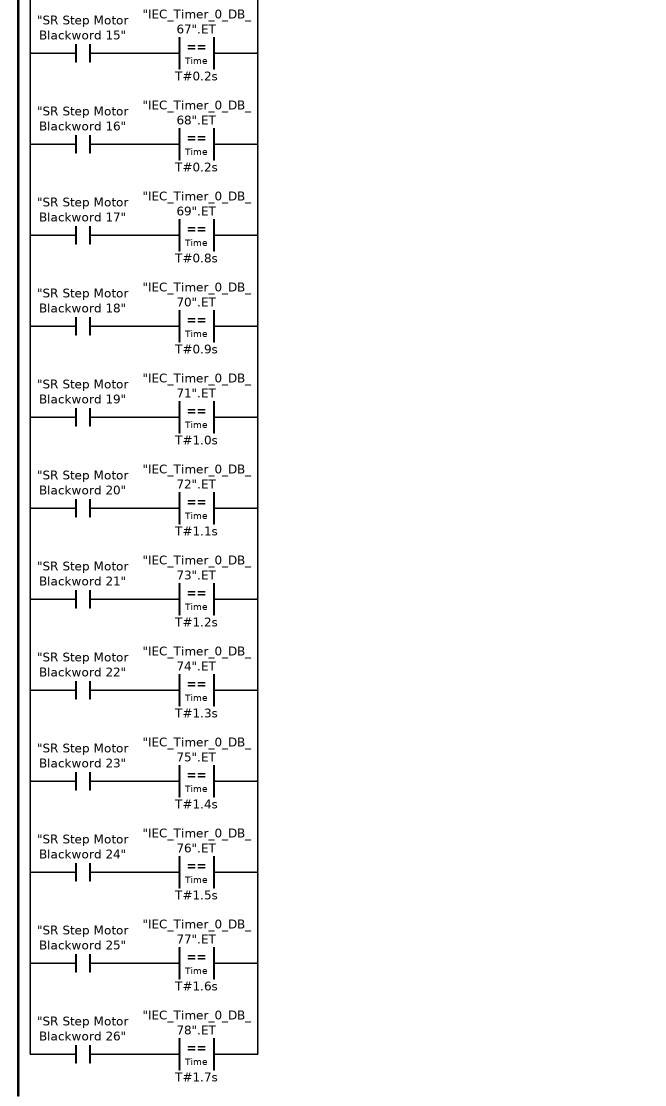
   "IEC_Counter_0_DB_1072".CTU(CU := ("SR Step Motor Blackword 1" AND ("IEC_Timer_0_DB_36".ET = T#2.0s)) OR ("SR Step Motor Blackword 2" AND ("IEC_Timer_0_DB_54".ET = T#1.9s)) OR ("SR Step Motor Blackword 3" AND ("IEC_Timer_0_DB_55".ET = T#1.8s)) OR ("SR Step Motor Blackword 4" AND ("IEC_Timer_0_DB_56".ET = T#1.7s)) OR ("SR Step Motor Blackword 5" AND ("IEC_Timer_0_DB_57".ET = T#1.6s)) OR ("SR Step Motor Blackword 6" AND ("IEC_Timer_0_DB_58".ET = T#1.5s)) OR ("SR Step Motor Blackword 7" AND ("IEC_Timer_0_DB_59".ET = T#1.4s)) OR ("SR Step Motor Blackword 8" AND ("IEC_Timer_0_DB_60".ET = T#1.3s)) OR ("SR Step Motor Blackword 9" AND ("IEC_Timer_0_DB_61".ET = T#1.2s)) OR ("SR Step Motor Blackword 10" AND ("IEC_Timer_0_DB_62".ET = T#1.1s)) OR ("SR Step Motor Blackword 11" AND ("IEC_Timer_0_DB_63".ET = T#1.0s)) OR ("SR Step Motor Blackword 12" AND ("IEC_Timer_0_DB_64".ET = T#0.9s)) OR ("SR Step Motor Blackword 13" AND ("IEC_Timer_0_DB_65".ET = T#0.8s)) OR ("SR Step Motor Blackword 14" AND ("IEC_Timer_0_DB_66".ET = T#0.2s)) OR ("SR Step Motor Blackword 15" AND ("IEC_Timer_0_DB_67".ET = T#0.2s)) OR ("SR Step Motor Blackword 16" AND ("IEC_Timer_0_DB_68".ET = T#0.2s)) OR ("SR Step Motor Blackword 17" AND ("IEC_Timer_0_DB_69".ET = T#0.8s)) OR ("SR Step Motor Blackword 18" AND ("IEC_Timer_0_DB_70".ET = T#0.9s)) OR ("SR Step Motor Blackword 19" AND ("IEC_Timer_0_DB_71".ET = T#1.0s)) OR ("SR Step Motor Blackword 20" AND ("IEC_Timer_0_DB_72".ET = T#1.1s)) OR ("SR Step Motor Blackword 21" AND ("IEC_Timer_0_DB_73".ET = T#1.2s)) OR ("SR Step Motor Blackword 22" AND ("IEC_Timer_0_DB_74".ET = T#1.3s)) OR ("SR Step Motor Blackword 23" AND ("IEC_Timer_0_DB_75".ET = T#1.4s)) OR ("SR Step Motor Blackword 24" AND ("IEC_Timer_0_DB_76".ET = T#1.5s)) OR ("SR Step Motor Blackword 25" AND ("IEC_Timer_0_DB_77".ET = T#1.6s)) OR ("SR Step Motor Blackword 26" AND ("IEC_Timer_0_DB_78".ET = T#1.7s)),
                           R := "Brushless Motor Conveyor ทำงาน",
                           PV := 1);
   "Output Reset พิเศษ จัดเก็บบ" := "IEC_Counter_0_DB_1072".Q;
END_REGION
END_FUNCTION_BLOCK

FUNCTION "Test" : Void   // FC5, LAD
{ S7_Optimized_Access := 'TRUE' }
VERSION : 0.1
BEGIN

REGION Network 1
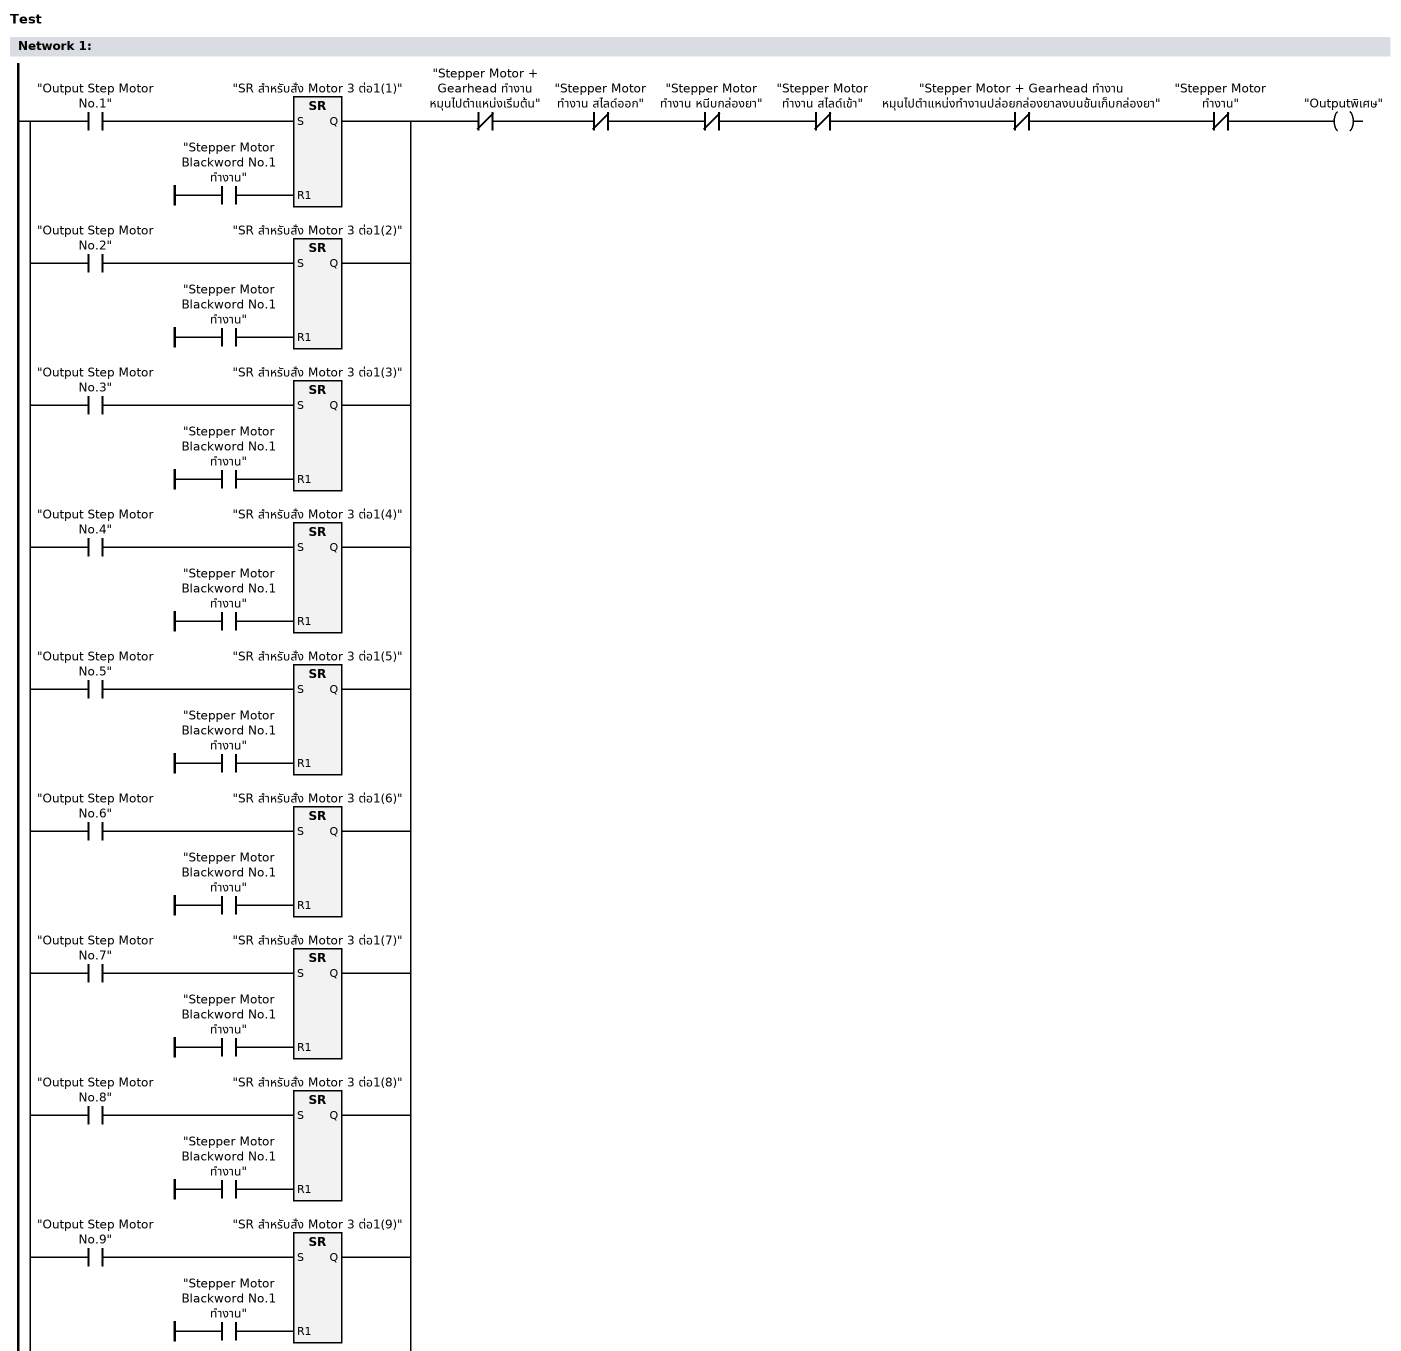
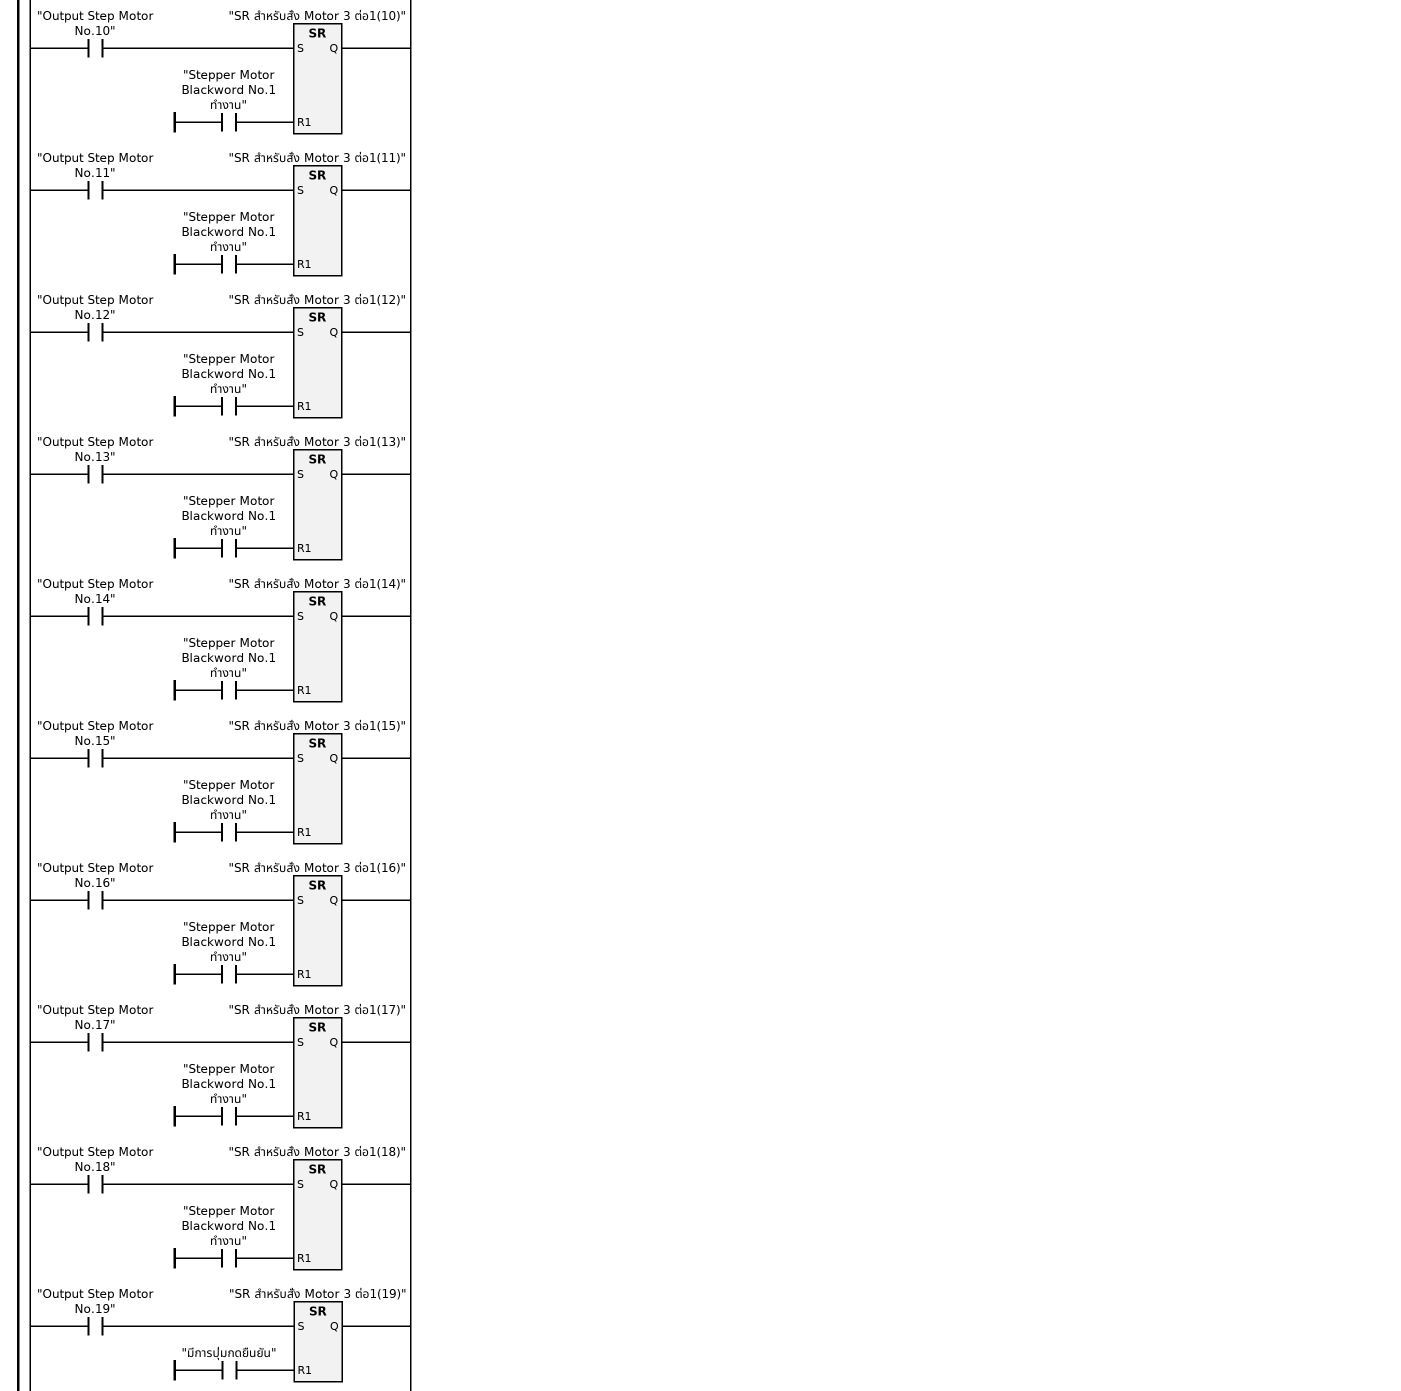
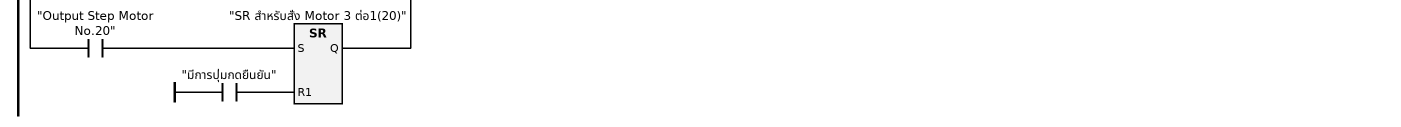
   RUNG wire#powerrail
      Contact( "Output Step Motor No.1" )
      S_SR(operand := "SR สำหรับสั่ง Motor 3 ต่อ1(1)", r1 := wire#w1)
      wire#w2
      I_Contact( "Stepper Motor + Gearhead ทำงาน หมุนไปตำแหน่งเริ่มต้น" )
      I_Contact( "Stepper Motor ทำงาน สไลด์ออก" )
      I_Contact( "Stepper Motor ทำงาน หนีบกล่องยา" )
      I_Contact( "Stepper Motor ทำงาน สไลด์เข้า" )
      I_Contact( "Stepper Motor + Gearhead ทำงาน หมุนไปตำแหน่งทำงานปล่อยกล่องยาลงบนชั้นเก็บกล่องยา" )
      I_Contact( "Stepper Motor  ทำงาน" )
      Coil( "Outputพิเศษ" )
   END_RUNG
   RUNG wire#powerrail
      Contact( "Stepper Motor Blackword No.1 ทำงาน" )
   END_RUNG wire#w1
   RUNG wire#powerrail
      Contact( "Output Step Motor No.2" )
      S_SR(operand := "SR สำหรับสั่ง Motor 3 ต่อ1(2)", r1 := wire#w3)
   END_RUNG wire#w2
   RUNG wire#powerrail
      Contact( "Stepper Motor Blackword No.1 ทำงาน" )
   END_RUNG wire#w3
   RUNG wire#powerrail
      Contact( "Output Step Motor No.3" )
      S_SR(operand := "SR สำหรับสั่ง Motor 3 ต่อ1(3)", r1 := wire#w4)
   END_RUNG wire#w2
   RUNG wire#powerrail
      Contact( "Stepper Motor Blackword No.1 ทำงาน" )
   END_RUNG wire#w4
   RUNG wire#powerrail
      Contact( "Output Step Motor No.4" )
      S_SR(operand := "SR สำหรับสั่ง Motor 3 ต่อ1(4)", r1 := wire#w5)
   END_RUNG wire#w2
   RUNG wire#powerrail
      Contact( "Stepper Motor Blackword No.1 ทำงาน" )
   END_RUNG wire#w5
   RUNG wire#powerrail
      Contact( "Output Step Motor No.5" )
      S_SR(operand := "SR สำหรับสั่ง Motor 3 ต่อ1(5)", r1 := wire#w6)
   END_RUNG wire#w2
   RUNG wire#powerrail
      Contact( "Stepper Motor Blackword No.1 ทำงาน" )
   END_RUNG wire#w6
   RUNG wire#powerrail
      Contact( "Output Step Motor No.6" )
      S_SR(operand := "SR สำหรับสั่ง Motor 3 ต่อ1(6)", r1 := wire#w7)
   END_RUNG wire#w2
   RUNG wire#powerrail
      Contact( "Stepper Motor Blackword No.1 ทำงาน" )
   END_RUNG wire#w7
   RUNG wire#powerrail
      Contact( "Output Step Motor No.7" )
      S_SR(operand := "SR สำหรับสั่ง Motor 3 ต่อ1(7)", r1 := wire#w8)
   END_RUNG wire#w2
   RUNG wire#powerrail
      Contact( "Stepper Motor Blackword No.1 ทำงาน" )
   END_RUNG wire#w8
   RUNG wire#powerrail
      Contact( "Output Step Motor No.8" )
      S_SR(operand := "SR สำหรับสั่ง Motor 3 ต่อ1(8)", r1 := wire#w9)
   END_RUNG wire#w2
   RUNG wire#powerrail
      Contact( "Stepper Motor Blackword No.1 ทำงาน" )
   END_RUNG wire#w9
   RUNG wire#powerrail
      Contact( "Output Step Motor No.9" )
      S_SR(operand := "SR สำหรับสั่ง Motor 3 ต่อ1(9)", r1 := wire#w10)
   END_RUNG wire#w2
   RUNG wire#powerrail
      Contact( "Stepper Motor Blackword No.1 ทำงาน" )
   END_RUNG wire#w10
   RUNG wire#powerrail
      Contact( "Output Step Motor No.10" )
      S_SR(operand := "SR สำหรับสั่ง Motor 3 ต่อ1(10)", r1 := wire#w11)
   END_RUNG wire#w2
   RUNG wire#powerrail
      Contact( "Stepper Motor Blackword No.1 ทำงาน" )
   END_RUNG wire#w11
   RUNG wire#powerrail
      Contact( "Output Step Motor No.11" )
      S_SR(operand := "SR สำหรับสั่ง Motor 3 ต่อ1(11)", r1 := wire#w12)
   END_RUNG wire#w2
   RUNG wire#powerrail
      Contact( "Stepper Motor Blackword No.1 ทำงาน" )
   END_RUNG wire#w12
   RUNG wire#powerrail
      Contact( "Output Step Motor No.12" )
      S_SR(operand := "SR สำหรับสั่ง Motor 3 ต่อ1(12)", r1 := wire#w13)
   END_RUNG wire#w2
   RUNG wire#powerrail
      Contact( "Stepper Motor Blackword No.1 ทำงาน" )
   END_RUNG wire#w13
   RUNG wire#powerrail
      Contact( "Output Step Motor No.13" )
      S_SR(operand := "SR สำหรับสั่ง Motor 3 ต่อ1(13)", r1 := wire#w14)
   END_RUNG wire#w2
   RUNG wire#powerrail
      Contact( "Stepper Motor Blackword No.1 ทำงาน" )
   END_RUNG wire#w14
   RUNG wire#powerrail
      Contact( "Output Step Motor No.14" )
      S_SR(operand := "SR สำหรับสั่ง Motor 3 ต่อ1(14)", r1 := wire#w15)
   END_RUNG wire#w2
   RUNG wire#powerrail
      Contact( "Stepper Motor Blackword No.1 ทำงาน" )
   END_RUNG wire#w15
   RUNG wire#powerrail
      Contact( "Output Step Motor No.15" )
      S_SR(operand := "SR สำหรับสั่ง Motor 3 ต่อ1(15)", r1 := wire#w16)
   END_RUNG wire#w2
   RUNG wire#powerrail
      Contact( "Stepper Motor Blackword No.1 ทำงาน" )
   END_RUNG wire#w16
   RUNG wire#powerrail
      Contact( "Output Step Motor No.16" )
      S_SR(operand := "SR สำหรับสั่ง Motor 3 ต่อ1(16)", r1 := wire#w17)
   END_RUNG wire#w2
   RUNG wire#powerrail
      Contact( "Stepper Motor Blackword No.1 ทำงาน" )
   END_RUNG wire#w17
   RUNG wire#powerrail
      Contact( "Output Step Motor No.17" )
      S_SR(operand := "SR สำหรับสั่ง Motor 3 ต่อ1(17)", r1 := wire#w18)
   END_RUNG wire#w2
   RUNG wire#powerrail
      Contact( "Stepper Motor Blackword No.1 ทำงาน" )
   END_RUNG wire#w18
   RUNG wire#powerrail
      Contact( "Output Step Motor No.18" )
      S_SR(operand := "SR สำหรับสั่ง Motor 3 ต่อ1(18)", r1 := wire#w19)
   END_RUNG wire#w2
   RUNG wire#powerrail
      Contact( "Stepper Motor Blackword No.1 ทำงาน" )
   END_RUNG wire#w19
   RUNG wire#powerrail
      Contact( "Output Step Motor No.19" )
      S_SR(operand := "SR สำหรับสั่ง Motor 3 ต่อ1(19)", r1 := wire#w20)
   END_RUNG wire#w2
   RUNG wire#powerrail
      Contact( "มีการปุ่มกดยืนยัน" )
   END_RUNG wire#w20
   RUNG wire#powerrail
      Contact( "Output Step Motor No.20" )
      S_SR(operand := "SR สำหรับสั่ง Motor 3 ต่อ1(20)", r1 := wire#w21)
   END_RUNG wire#w2
   RUNG wire#powerrail
      Contact( "มีการปุ่มกดยืนยัน" )
   END_RUNG wire#w21
   // the same network as SCL:
   IF "Output Step Motor No.1" THEN
       "SR สำหรับสั่ง Motor 3 ต่อ1(1)" := TRUE;   // SR flip-flop
   END_IF;
   IF "Stepper Motor Blackword No.1 ทำงาน" THEN "SR สำหรับสั่ง Motor 3 ต่อ1(1)" := FALSE; END_IF;
   IF "Output Step Motor No.2" THEN
       "SR สำหรับสั่ง Motor 3 ต่อ1(2)" := TRUE;   // SR flip-flop
   END_IF;
   IF "Stepper Motor Blackword No.1 ทำงาน" THEN "SR สำหรับสั่ง Motor 3 ต่อ1(2)" := FALSE; END_IF;
   IF "Output Step Motor No.3" THEN
       "SR สำหรับสั่ง Motor 3 ต่อ1(3)" := TRUE;   // SR flip-flop
   END_IF;
   IF "Stepper Motor Blackword No.1 ทำงาน" THEN "SR สำหรับสั่ง Motor 3 ต่อ1(3)" := FALSE; END_IF;
   IF "Output Step Motor No.4" THEN
       "SR สำหรับสั่ง Motor 3 ต่อ1(4)" := TRUE;   // SR flip-flop
   END_IF;
   IF "Stepper Motor Blackword No.1 ทำงาน" THEN "SR สำหรับสั่ง Motor 3 ต่อ1(4)" := FALSE; END_IF;
   IF "Output Step Motor No.5" THEN
       "SR สำหรับสั่ง Motor 3 ต่อ1(5)" := TRUE;   // SR flip-flop
   END_IF;
   IF "Stepper Motor Blackword No.1 ทำงาน" THEN "SR สำหรับสั่ง Motor 3 ต่อ1(5)" := FALSE; END_IF;
   IF "Output Step Motor No.6" THEN
       "SR สำหรับสั่ง Motor 3 ต่อ1(6)" := TRUE;   // SR flip-flop
   END_IF;
   IF "Stepper Motor Blackword No.1 ทำงาน" THEN "SR สำหรับสั่ง Motor 3 ต่อ1(6)" := FALSE; END_IF;
   IF "Output Step Motor No.7" THEN
       "SR สำหรับสั่ง Motor 3 ต่อ1(7)" := TRUE;   // SR flip-flop
   END_IF;
   IF "Stepper Motor Blackword No.1 ทำงาน" THEN "SR สำหรับสั่ง Motor 3 ต่อ1(7)" := FALSE; END_IF;
   IF "Output Step Motor No.8" THEN
       "SR สำหรับสั่ง Motor 3 ต่อ1(8)" := TRUE;   // SR flip-flop
   END_IF;
   IF "Stepper Motor Blackword No.1 ทำงาน" THEN "SR สำหรับสั่ง Motor 3 ต่อ1(8)" := FALSE; END_IF;
   IF "Output Step Motor No.9" THEN
       "SR สำหรับสั่ง Motor 3 ต่อ1(9)" := TRUE;   // SR flip-flop
   END_IF;
   IF "Stepper Motor Blackword No.1 ทำงาน" THEN "SR สำหรับสั่ง Motor 3 ต่อ1(9)" := FALSE; END_IF;
   IF "Output Step Motor No.10" THEN
       "SR สำหรับสั่ง Motor 3 ต่อ1(10)" := TRUE;   // SR flip-flop
   END_IF;
   IF "Stepper Motor Blackword No.1 ทำงาน" THEN "SR สำหรับสั่ง Motor 3 ต่อ1(10)" := FALSE; END_IF;
   IF "Output Step Motor No.11" THEN
       "SR สำหรับสั่ง Motor 3 ต่อ1(11)" := TRUE;   // SR flip-flop
   END_IF;
   IF "Stepper Motor Blackword No.1 ทำงาน" THEN "SR สำหรับสั่ง Motor 3 ต่อ1(11)" := FALSE; END_IF;
   IF "Output Step Motor No.12" THEN
       "SR สำหรับสั่ง Motor 3 ต่อ1(12)" := TRUE;   // SR flip-flop
   END_IF;
   IF "Stepper Motor Blackword No.1 ทำงาน" THEN "SR สำหรับสั่ง Motor 3 ต่อ1(12)" := FALSE; END_IF;
   IF "Output Step Motor No.13" THEN
       "SR สำหรับสั่ง Motor 3 ต่อ1(13)" := TRUE;   // SR flip-flop
   END_IF;
   IF "Stepper Motor Blackword No.1 ทำงาน" THEN "SR สำหรับสั่ง Motor 3 ต่อ1(13)" := FALSE; END_IF;
   IF "Output Step Motor No.14" THEN
       "SR สำหรับสั่ง Motor 3 ต่อ1(14)" := TRUE;   // SR flip-flop
   END_IF;
   IF "Stepper Motor Blackword No.1 ทำงาน" THEN "SR สำหรับสั่ง Motor 3 ต่อ1(14)" := FALSE; END_IF;
   IF "Output Step Motor No.15" THEN
       "SR สำหรับสั่ง Motor 3 ต่อ1(15)" := TRUE;   // SR flip-flop
   END_IF;
   IF "Stepper Motor Blackword No.1 ทำงาน" THEN "SR สำหรับสั่ง Motor 3 ต่อ1(15)" := FALSE; END_IF;
   IF "Output Step Motor No.16" THEN
       "SR สำหรับสั่ง Motor 3 ต่อ1(16)" := TRUE;   // SR flip-flop
   END_IF;
   IF "Stepper Motor Blackword No.1 ทำงาน" THEN "SR สำหรับสั่ง Motor 3 ต่อ1(16)" := FALSE; END_IF;
   IF "Output Step Motor No.17" THEN
       "SR สำหรับสั่ง Motor 3 ต่อ1(17)" := TRUE;   // SR flip-flop
   END_IF;
   IF "Stepper Motor Blackword No.1 ทำงาน" THEN "SR สำหรับสั่ง Motor 3 ต่อ1(17)" := FALSE; END_IF;
   IF "Output Step Motor No.18" THEN
       "SR สำหรับสั่ง Motor 3 ต่อ1(18)" := TRUE;   // SR flip-flop
   END_IF;
   IF "Stepper Motor Blackword No.1 ทำงาน" THEN "SR สำหรับสั่ง Motor 3 ต่อ1(18)" := FALSE; END_IF;
   IF "Output Step Motor No.19" THEN
       "SR สำหรับสั่ง Motor 3 ต่อ1(19)" := TRUE;   // SR flip-flop
   END_IF;
   IF "มีการปุ่มกดยืนยัน" THEN "SR สำหรับสั่ง Motor 3 ต่อ1(19)" := FALSE; END_IF;
   IF "Output Step Motor No.20" THEN
       "SR สำหรับสั่ง Motor 3 ต่อ1(20)" := TRUE;   // SR flip-flop
   END_IF;
   IF "มีการปุ่มกดยืนยัน" THEN "SR สำหรับสั่ง Motor 3 ต่อ1(20)" := FALSE; END_IF;
   "Outputพิเศษ" := ("SR สำหรับสั่ง Motor 3 ต่อ1(1)" OR "SR สำหรับสั่ง Motor 3 ต่อ1(2)" OR "SR สำหรับสั่ง Motor 3 ต่อ1(3)" OR "SR สำหรับสั่ง Motor 3 ต่อ1(4)" OR "SR สำหรับสั่ง Motor 3 ต่อ1(5)" OR "SR สำหรับสั่ง Motor 3 ต่อ1(6)" OR "SR สำหรับสั่ง Motor 3 ต่อ1(7)" OR "SR สำหรับสั่ง Motor 3 ต่อ1(8)" OR "SR สำหรับสั่ง Motor 3 ต่อ1(9)" OR "SR สำหรับสั่ง Motor 3 ต่อ1(10)" OR "SR สำหรับสั่ง Motor 3 ต่อ1(11)" OR "SR สำหรับสั่ง Motor 3 ต่อ1(12)" OR "SR สำหรับสั่ง Motor 3 ต่อ1(13)" OR "SR สำหรับสั่ง Motor 3 ต่อ1(14)" OR "SR สำหรับสั่ง Motor 3 ต่อ1(15)" OR "SR สำหรับสั่ง Motor 3 ต่อ1(16)" OR "SR สำหรับสั่ง Motor 3 ต่อ1(17)" OR "SR สำหรับสั่ง Motor 3 ต่อ1(18)" OR "SR สำหรับสั่ง Motor 3 ต่อ1(19)" OR "SR สำหรับสั่ง Motor 3 ต่อ1(20)") AND NOT "Stepper Motor + Gearhead ทำงาน หมุนไปตำแหน่งเริ่มต้น" AND NOT "Stepper Motor ทำงาน สไลด์ออก" AND NOT "Stepper Motor ทำงาน หนีบกล่องยา" AND NOT "Stepper Motor ทำงาน สไลด์เข้า" AND NOT "Stepper Motor + Gearhead ทำงาน หมุนไปตำแหน่งทำงานปล่อยกล่องยาลงบนชั้นเก็บกล่องยา" AND NOT "Stepper Motor  ทำงาน";
END_REGION
END_FUNCTION

FUNCTION "Test1" : Void   // FC9, LAD
{ S7_Optimized_Access := 'TRUE' }
VERSION : 0.1
   VAR_OUTPUT
      "Output  (พิเศษ)" : Bool;
   END_VAR
BEGIN

REGION Network 1
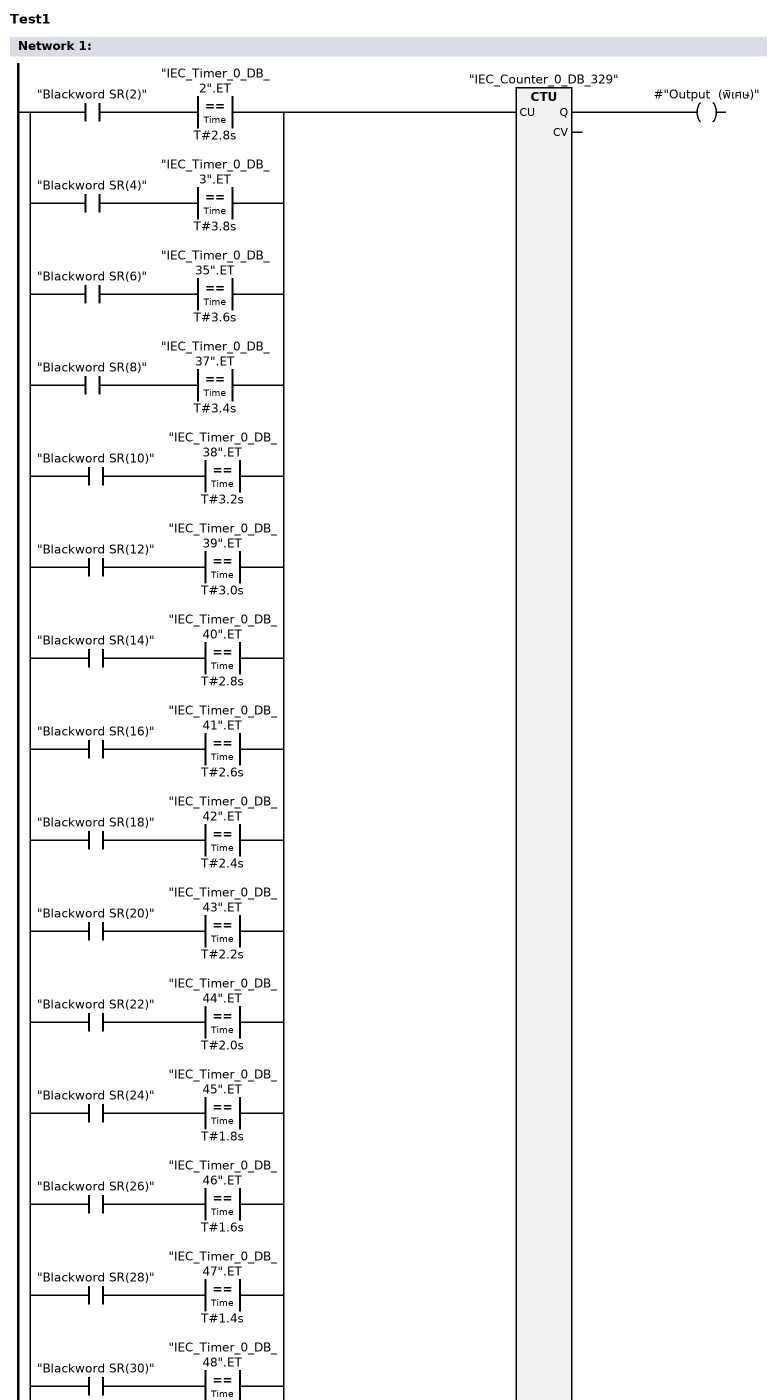
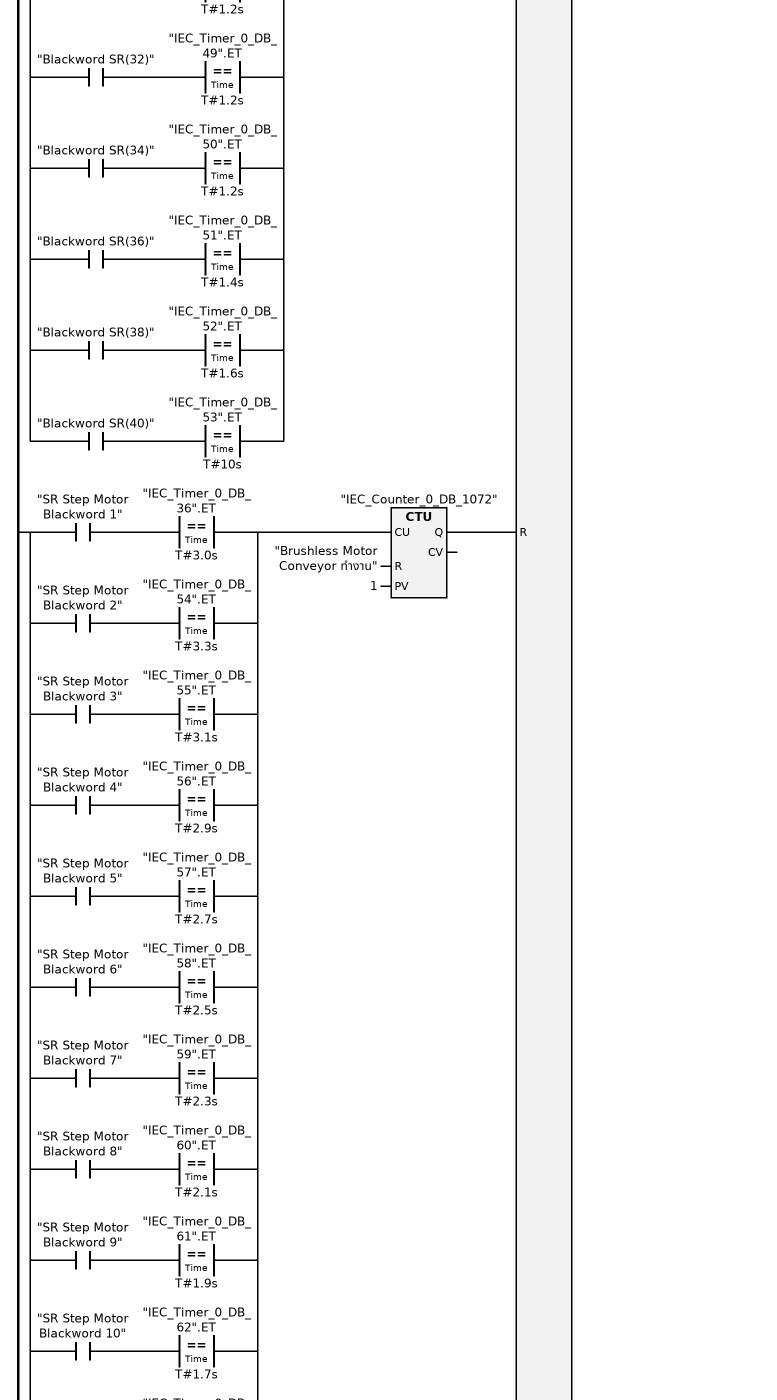
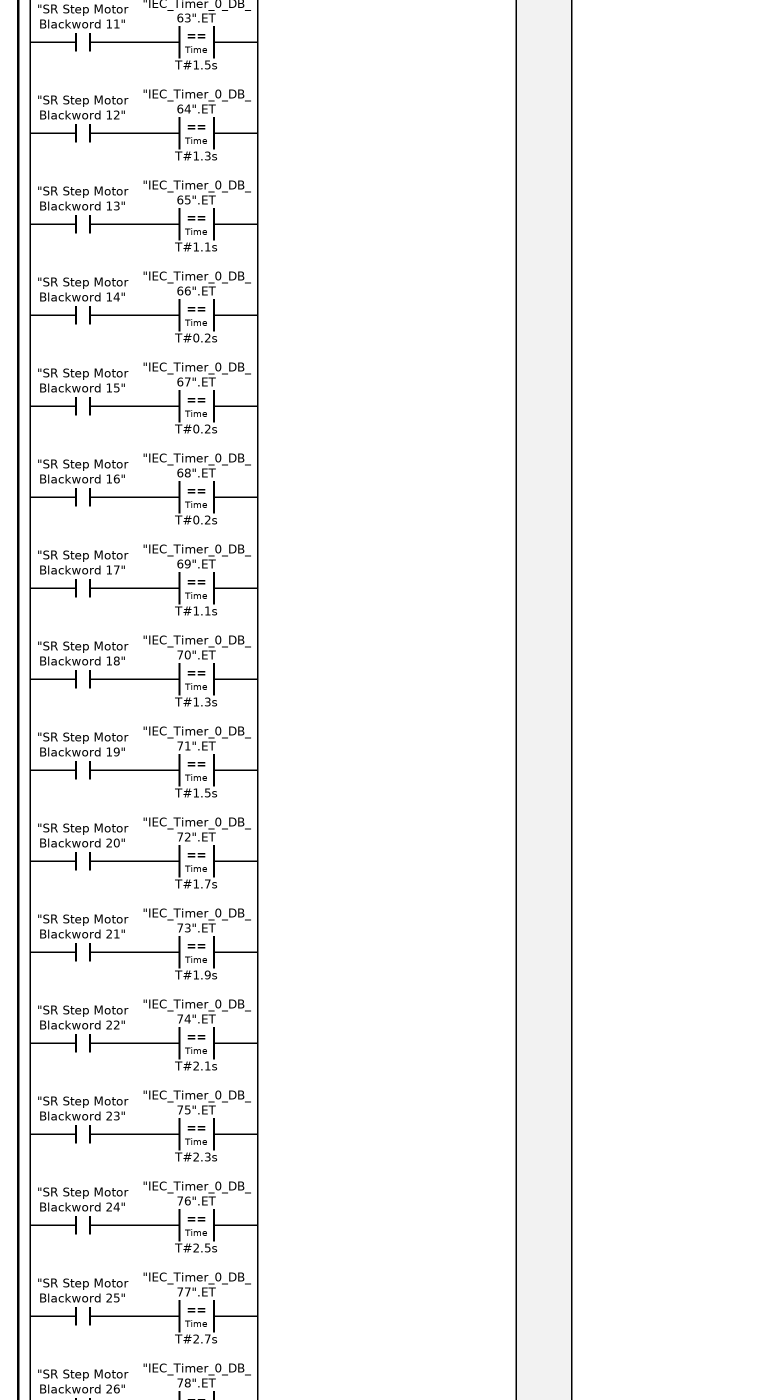
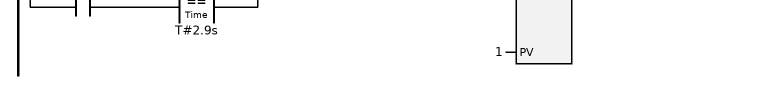
   "IEC_Counter_0_DB_1072".CTU(CU := ("SR Step Motor Blackword 1" AND ("IEC_Timer_0_DB_36".ET = T#3.0s)) OR ("SR Step Motor Blackword 2" AND ("IEC_Timer_0_DB_54".ET = T#3.3s)) OR ("SR Step Motor Blackword 3" AND ("IEC_Timer_0_DB_55".ET = T#3.1s)) OR ("SR Step Motor Blackword 4" AND ("IEC_Timer_0_DB_56".ET = T#2.9s)) OR ("SR Step Motor Blackword 5" AND ("IEC_Timer_0_DB_57".ET = T#2.7s)) OR ("SR Step Motor Blackword 6" AND ("IEC_Timer_0_DB_58".ET = T#2.5s)) OR ("SR Step Motor Blackword 7" AND ("IEC_Timer_0_DB_59".ET = T#2.3s)) OR ("SR Step Motor Blackword 8" AND ("IEC_Timer_0_DB_60".ET = T#2.1s)) OR ("SR Step Motor Blackword 9" AND ("IEC_Timer_0_DB_61".ET = T#1.9s)) OR ("SR Step Motor Blackword 10" AND ("IEC_Timer_0_DB_62".ET = T#1.7s)) OR ("SR Step Motor Blackword 11" AND ("IEC_Timer_0_DB_63".ET = T#1.5s)) OR ("SR Step Motor Blackword 12" AND ("IEC_Timer_0_DB_64".ET = T#1.3s)) OR ("SR Step Motor Blackword 13" AND ("IEC_Timer_0_DB_65".ET = T#1.1s)) OR ("SR Step Motor Blackword 14" AND ("IEC_Timer_0_DB_66".ET = T#0.2s)) OR ("SR Step Motor Blackword 15" AND ("IEC_Timer_0_DB_67".ET = T#0.2s)) OR ("SR Step Motor Blackword 16" AND ("IEC_Timer_0_DB_68".ET = T#0.2s)) OR ("SR Step Motor Blackword 17" AND ("IEC_Timer_0_DB_69".ET = T#1.1s)) OR ("SR Step Motor Blackword 18" AND ("IEC_Timer_0_DB_70".ET = T#1.3s)) OR ("SR Step Motor Blackword 19" AND ("IEC_Timer_0_DB_71".ET = T#1.5s)) OR ("SR Step Motor Blackword 20" AND ("IEC_Timer_0_DB_72".ET = T#1.7s)) OR ("SR Step Motor Blackword 21" AND ("IEC_Timer_0_DB_73".ET = T#1.9s)) OR ("SR Step Motor Blackword 22" AND ("IEC_Timer_0_DB_74".ET = T#2.1s)) OR ("SR Step Motor Blackword 23" AND ("IEC_Timer_0_DB_75".ET = T#2.3s)) OR ("SR Step Motor Blackword 24" AND ("IEC_Timer_0_DB_76".ET = T#2.5s)) OR ("SR Step Motor Blackword 25" AND ("IEC_Timer_0_DB_77".ET = T#2.7s)) OR ("SR Step Motor Blackword 26" AND ("IEC_Timer_0_DB_78".ET = T#2.9s)),
                           R := "Brushless Motor Conveyor ทำงาน",
                           PV := 1);
   "IEC_Counter_0_DB_329".CTU(CU := ("Blackword SR(2)" AND ("IEC_Timer_0_DB_2".ET = T#2.8s)) OR ("Blackword SR(4)" AND ("IEC_Timer_0_DB_3".ET = T#3.8s)) OR ("Blackword SR(6)" AND ("IEC_Timer_0_DB_35".ET = T#3.6s)) OR ("Blackword SR(8)" AND ("IEC_Timer_0_DB_37".ET = T#3.4s)) OR ("Blackword SR(10)" AND ("IEC_Timer_0_DB_38".ET = T#3.2s)) OR ("Blackword SR(12)" AND ("IEC_Timer_0_DB_39".ET = T#3.0s)) OR ("Blackword SR(14)" AND ("IEC_Timer_0_DB_40".ET = T#2.8s)) OR ("Blackword SR(16)" AND ("IEC_Timer_0_DB_41".ET = T#2.6s)) OR ("Blackword SR(18)" AND ("IEC_Timer_0_DB_42".ET = T#2.4s)) OR ("Blackword SR(20)" AND ("IEC_Timer_0_DB_43".ET = T#2.2s)) OR ("Blackword SR(22)" AND ("IEC_Timer_0_DB_44".ET = T#2.0s)) OR ("Blackword SR(24)" AND ("IEC_Timer_0_DB_45".ET = T#1.8s)) OR ("Blackword SR(26)" AND ("IEC_Timer_0_DB_46".ET = T#1.6s)) OR ("Blackword SR(28)" AND ("IEC_Timer_0_DB_47".ET = T#1.4s)) OR ("Blackword SR(30)" AND ("IEC_Timer_0_DB_48".ET = T#1.2s)) OR ("Blackword SR(32)" AND ("IEC_Timer_0_DB_49".ET = T#1.2s)) OR ("Blackword SR(34)" AND ("IEC_Timer_0_DB_50".ET = T#1.2s)) OR ("Blackword SR(36)" AND ("IEC_Timer_0_DB_51".ET = T#1.4s)) OR ("Blackword SR(38)" AND ("IEC_Timer_0_DB_52".ET = T#1.6s)) OR ("Blackword SR(40)" AND ("IEC_Timer_0_DB_53".ET = T#10s)),
                           R := "IEC_Counter_0_DB_1072".Q,
                           PV := 1);
   #"Output  (พิเศษ)" := "IEC_Counter_0_DB_329".Q;
END_REGION
END_FUNCTION

// folder: System_Out(เบิกจ่าย)

FUNCTION "ตัวเลือกยา (26)" : Void   // FC8, LAD
{ S7_Optimized_Access := 'TRUE' }
VERSION : 0.1
   VAR_INPUT
      "ปึ่ม 1" : Int;
      "ปึ่ม 2" : Int;
      "ปึ่ม 3" : Int;
      "ปึ่ม 4" : Int;
      "ปึ่ม 5" : Int;
      "ปึ่ม 6" : Int;
      "ปึ่ม 7" : Int;
      "ปึ่ม 8" : Int;
      "ปึ่ม 9" : Int;
      "ปึ่ม 10" : Int;
      "ปึ่ม 11" : Int;
      "ปึ่ม 12" : Int;
      "ปึ่ม 13" : Int;
      "ปึ่ม 14" : Int;
      "ปึ่ม 15" : Int;
      "ปึ่ม 16" : Int;
      "ปึ่ม 17" : Int;
      "ปึ่ม 18" : Int;
      "ปึ่ม 19" : Int;
      "ปึ่ม 20" : Int;
      "ปึ่ม 21" : Int;
      "ปึ่ม 22" : Int;
      "ปึ่ม 23" : Int;
      "ปึ่ม 24" : Int;
      "ปึ่ม 25" : Int;
      "ปึ่ม 26" : Int;
   END_VAR
   VAR_OUTPUT
      "เมื่ิอมีการกดปุ้ม" : Bool;
   END_VAR
BEGIN

REGION Network 1
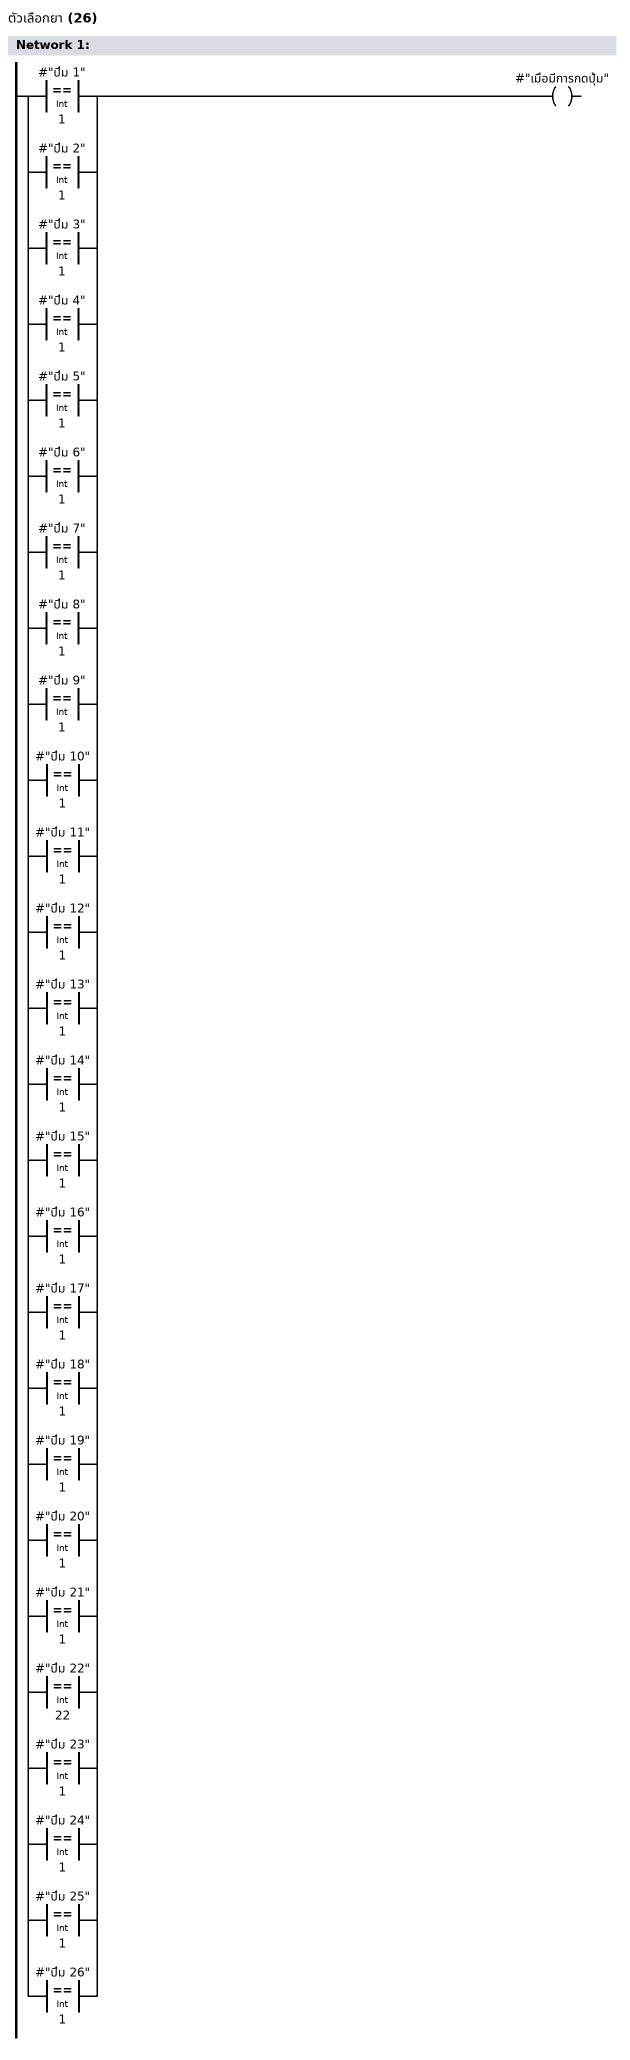
   RUNG wire#powerrail
      { S7_Templates := "SrcType := Int" } EQ_Contact(in1 := #"ปึ่ม 1", in2 := 1)
      wire#w1
      Coil( #"เมื่ิอมีการกดปุ้ม" )
   END_RUNG
   RUNG wire#powerrail
      { S7_Templates := "SrcType := Int" } EQ_Contact(in1 := #"ปึ่ม 2", in2 := 1)
   END_RUNG wire#w1
   RUNG wire#powerrail
      { S7_Templates := "SrcType := Int" } EQ_Contact(in1 := #"ปึ่ม 3", in2 := 1)
   END_RUNG wire#w1
   RUNG wire#powerrail
      { S7_Templates := "SrcType := Int" } EQ_Contact(in1 := #"ปึ่ม 4", in2 := 1)
   END_RUNG wire#w1
   RUNG wire#powerrail
      { S7_Templates := "SrcType := Int" } EQ_Contact(in1 := #"ปึ่ม 5", in2 := 1)
   END_RUNG wire#w1
   RUNG wire#powerrail
      { S7_Templates := "SrcType := Int" } EQ_Contact(in1 := #"ปึ่ม 6", in2 := 1)
   END_RUNG wire#w1
   RUNG wire#powerrail
      { S7_Templates := "SrcType := Int" } EQ_Contact(in1 := #"ปึ่ม 7", in2 := 1)
   END_RUNG wire#w1
   RUNG wire#powerrail
      { S7_Templates := "SrcType := Int" } EQ_Contact(in1 := #"ปึ่ม 8", in2 := 1)
   END_RUNG wire#w1
   RUNG wire#powerrail
      { S7_Templates := "SrcType := Int" } EQ_Contact(in1 := #"ปึ่ม 9", in2 := 1)
   END_RUNG wire#w1
   RUNG wire#powerrail
      { S7_Templates := "SrcType := Int" } EQ_Contact(in1 := #"ปึ่ม 10", in2 := 1)
   END_RUNG wire#w1
   RUNG wire#powerrail
      { S7_Templates := "SrcType := Int" } EQ_Contact(in1 := #"ปึ่ม 11", in2 := 1)
   END_RUNG wire#w1
   RUNG wire#powerrail
      { S7_Templates := "SrcType := Int" } EQ_Contact(in1 := #"ปึ่ม 12", in2 := 1)
   END_RUNG wire#w1
   RUNG wire#powerrail
      { S7_Templates := "SrcType := Int" } EQ_Contact(in1 := #"ปึ่ม 13", in2 := 1)
   END_RUNG wire#w1
   RUNG wire#powerrail
      { S7_Templates := "SrcType := Int" } EQ_Contact(in1 := #"ปึ่ม 14", in2 := 1)
   END_RUNG wire#w1
   RUNG wire#powerrail
      { S7_Templates := "SrcType := Int" } EQ_Contact(in1 := #"ปึ่ม 15", in2 := 1)
   END_RUNG wire#w1
   RUNG wire#powerrail
      { S7_Templates := "SrcType := Int" } EQ_Contact(in1 := #"ปึ่ม 16", in2 := 1)
   END_RUNG wire#w1
   RUNG wire#powerrail
      { S7_Templates := "SrcType := Int" } EQ_Contact(in1 := #"ปึ่ม 17", in2 := 1)
   END_RUNG wire#w1
   RUNG wire#powerrail
      { S7_Templates := "SrcType := Int" } EQ_Contact(in1 := #"ปึ่ม 18", in2 := 1)
   END_RUNG wire#w1
   RUNG wire#powerrail
      { S7_Templates := "SrcType := Int" } EQ_Contact(in1 := #"ปึ่ม 19", in2 := 1)
   END_RUNG wire#w1
   RUNG wire#powerrail
      { S7_Templates := "SrcType := Int" } EQ_Contact(in1 := #"ปึ่ม 20", in2 := 1)
   END_RUNG wire#w1
   RUNG wire#powerrail
      { S7_Templates := "SrcType := Int" } EQ_Contact(in1 := #"ปึ่ม 21", in2 := 1)
   END_RUNG wire#w1
   RUNG wire#powerrail
      { S7_Templates := "SrcType := Int" } EQ_Contact(in1 := #"ปึ่ม 22", in2 := 22)
   END_RUNG wire#w1
   RUNG wire#powerrail
      { S7_Templates := "SrcType := Int" } EQ_Contact(in1 := #"ปึ่ม 23", in2 := 1)
   END_RUNG wire#w1
   RUNG wire#powerrail
      { S7_Templates := "SrcType := Int" } EQ_Contact(in1 := #"ปึ่ม 24", in2 := 1)
   END_RUNG wire#w1
   RUNG wire#powerrail
      { S7_Templates := "SrcType := Int" } EQ_Contact(in1 := #"ปึ่ม 25", in2 := 1)
   END_RUNG wire#w1
   RUNG wire#powerrail
      { S7_Templates := "SrcType := Int" } EQ_Contact(in1 := #"ปึ่ม 26", in2 := 1)
   END_RUNG wire#w1
   // the same network as SCL:
   #"เมื่ิอมีการกดปุ้ม" := (#"ปึ่ม 1" = 1) OR (#"ปึ่ม 2" = 1) OR (#"ปึ่ม 3" = 1) OR (#"ปึ่ม 4" = 1) OR (#"ปึ่ม 5" = 1) OR (#"ปึ่ม 6" = 1) OR (#"ปึ่ม 7" = 1) OR (#"ปึ่ม 8" = 1) OR (#"ปึ่ม 9" = 1) OR (#"ปึ่ม 10" = 1) OR (#"ปึ่ม 11" = 1) OR (#"ปึ่ม 12" = 1) OR (#"ปึ่ม 13" = 1) OR (#"ปึ่ม 14" = 1) OR (#"ปึ่ม 15" = 1) OR (#"ปึ่ม 16" = 1) OR (#"ปึ่ม 17" = 1) OR (#"ปึ่ม 18" = 1) OR (#"ปึ่ม 19" = 1) OR (#"ปึ่ม 20" = 1) OR (#"ปึ่ม 21" = 1) OR (#"ปึ่ม 22" = 22) OR (#"ปึ่ม 23" = 1) OR (#"ปึ่ม 24" = 1) OR (#"ปึ่ม 25" = 1) OR (#"ปึ่ม 26" = 1);
END_REGION
END_FUNCTION

FUNCTION "ตัวเลือกยา (20)" : Void   // FC11, LAD
{ S7_Optimized_Access := 'TRUE' }
VERSION : 0.1
   VAR_INPUT
      "ปึ่ม 1" : Int;
      "ปึ่ม 2" : Int;
      "ปึ่ม 3" : Int;
      "ปึ่ม 4" : Int;
      "ปึ่ม 5" : Int;
      "ปึ่ม 6" : Int;
      "ปึ่ม 7" : Int;
      "ปึ่ม 8" : Int;
      "ปึ่ม 9" : Int;
      "ปึ่ม 10" : Int;
      "ปึ่ม 11" : Int;
      "ปึ่ม 12" : Int;
      "ปึ่ม 13" : Int;
      "ปึ่ม 14" : Int;
      "ปึ่ม 15" : Int;
      "ปึ่ม 16" : Int;
      "ปึ่ม 17" : Int;
      "ปึ่ม 18" : Int;
      "ปึ่ม 19" : Int;
      "ปึ่ม 20" : Int;
   END_VAR
   VAR_OUTPUT
      "เมื่อกดปุ่ม" : Bool;
   END_VAR
BEGIN

REGION Network 1
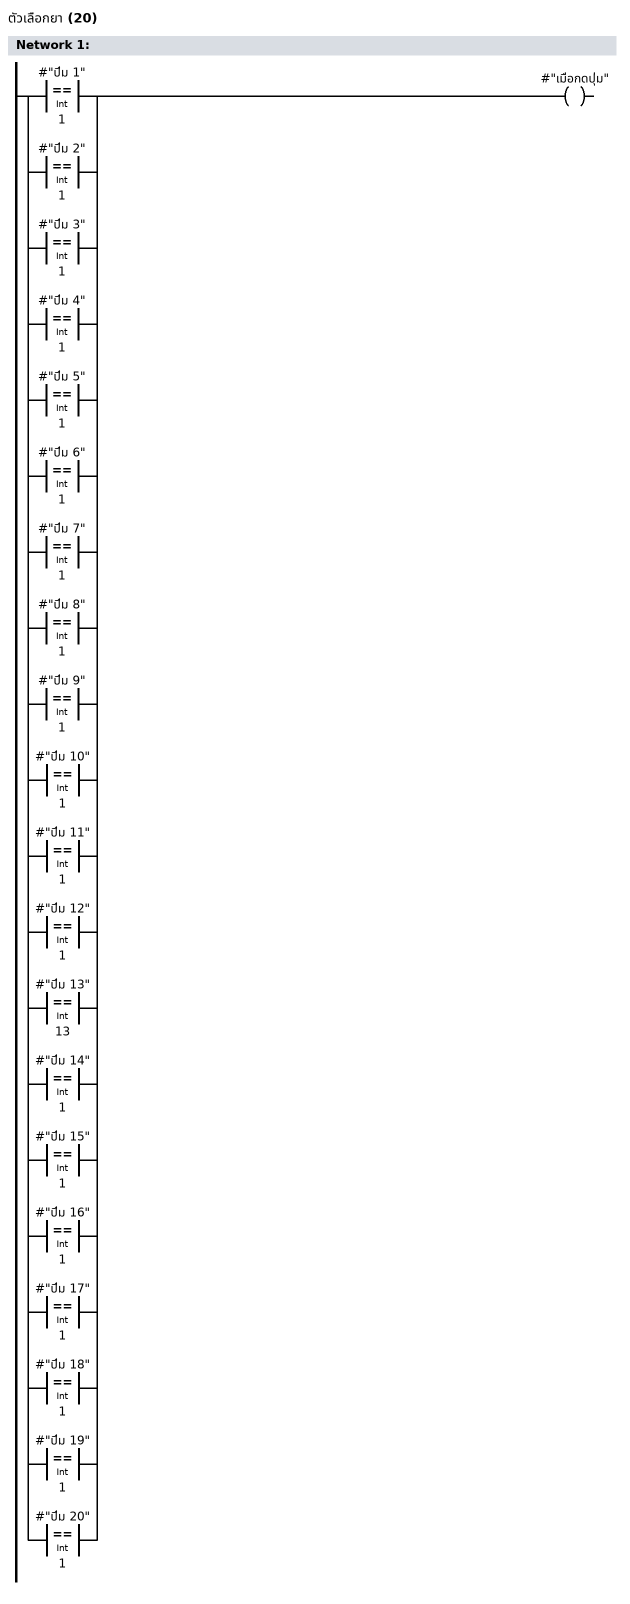
   RUNG wire#powerrail
      { S7_Templates := "SrcType := Int" } EQ_Contact(in1 := #"ปึ่ม 1", in2 := 1)
      wire#w1
      Coil( #"เมื่อกดปุ่ม" )
   END_RUNG
   RUNG wire#powerrail
      { S7_Templates := "SrcType := Int" } EQ_Contact(in1 := #"ปึ่ม 2", in2 := 1)
   END_RUNG wire#w1
   RUNG wire#powerrail
      { S7_Templates := "SrcType := Int" } EQ_Contact(in1 := #"ปึ่ม 3", in2 := 1)
   END_RUNG wire#w1
   RUNG wire#powerrail
      { S7_Templates := "SrcType := Int" } EQ_Contact(in1 := #"ปึ่ม 4", in2 := 1)
   END_RUNG wire#w1
   RUNG wire#powerrail
      { S7_Templates := "SrcType := Int" } EQ_Contact(in1 := #"ปึ่ม 5", in2 := 1)
   END_RUNG wire#w1
   RUNG wire#powerrail
      { S7_Templates := "SrcType := Int" } EQ_Contact(in1 := #"ปึ่ม 6", in2 := 1)
   END_RUNG wire#w1
   RUNG wire#powerrail
      { S7_Templates := "SrcType := Int" } EQ_Contact(in1 := #"ปึ่ม 7", in2 := 1)
   END_RUNG wire#w1
   RUNG wire#powerrail
      { S7_Templates := "SrcType := Int" } EQ_Contact(in1 := #"ปึ่ม 8", in2 := 1)
   END_RUNG wire#w1
   RUNG wire#powerrail
      { S7_Templates := "SrcType := Int" } EQ_Contact(in1 := #"ปึ่ม 9", in2 := 1)
   END_RUNG wire#w1
   RUNG wire#powerrail
      { S7_Templates := "SrcType := Int" } EQ_Contact(in1 := #"ปึ่ม 10", in2 := 1)
   END_RUNG wire#w1
   RUNG wire#powerrail
      { S7_Templates := "SrcType := Int" } EQ_Contact(in1 := #"ปึ่ม 11", in2 := 1)
   END_RUNG wire#w1
   RUNG wire#powerrail
      { S7_Templates := "SrcType := Int" } EQ_Contact(in1 := #"ปึ่ม 12", in2 := 1)
   END_RUNG wire#w1
   RUNG wire#powerrail
      { S7_Templates := "SrcType := Int" } EQ_Contact(in1 := #"ปึ่ม 13", in2 := 13)
   END_RUNG wire#w1
   RUNG wire#powerrail
      { S7_Templates := "SrcType := Int" } EQ_Contact(in1 := #"ปึ่ม 14", in2 := 1)
   END_RUNG wire#w1
   RUNG wire#powerrail
      { S7_Templates := "SrcType := Int" } EQ_Contact(in1 := #"ปึ่ม 15", in2 := 1)
   END_RUNG wire#w1
   RUNG wire#powerrail
      { S7_Templates := "SrcType := Int" } EQ_Contact(in1 := #"ปึ่ม 16", in2 := 1)
   END_RUNG wire#w1
   RUNG wire#powerrail
      { S7_Templates := "SrcType := Int" } EQ_Contact(in1 := #"ปึ่ม 17", in2 := 1)
   END_RUNG wire#w1
   RUNG wire#powerrail
      { S7_Templates := "SrcType := Int" } EQ_Contact(in1 := #"ปึ่ม 18", in2 := 1)
   END_RUNG wire#w1
   RUNG wire#powerrail
      { S7_Templates := "SrcType := Int" } EQ_Contact(in1 := #"ปึ่ม 19", in2 := 1)
   END_RUNG wire#w1
   RUNG wire#powerrail
      { S7_Templates := "SrcType := Int" } EQ_Contact(in1 := #"ปึ่ม 20", in2 := 1)
   END_RUNG wire#w1
   // the same network as SCL:
   #"เมื่อกดปุ่ม" := (#"ปึ่ม 1" = 1) OR (#"ปึ่ม 2" = 1) OR (#"ปึ่ม 3" = 1) OR (#"ปึ่ม 4" = 1) OR (#"ปึ่ม 5" = 1) OR (#"ปึ่ม 6" = 1) OR (#"ปึ่ม 7" = 1) OR (#"ปึ่ม 8" = 1) OR (#"ปึ่ม 9" = 1) OR (#"ปึ่ม 10" = 1) OR (#"ปึ่ม 11" = 1) OR (#"ปึ่ม 12" = 1) OR (#"ปึ่ม 13" = 13) OR (#"ปึ่ม 14" = 1) OR (#"ปึ่ม 15" = 1) OR (#"ปึ่ม 16" = 1) OR (#"ปึ่ม 17" = 1) OR (#"ปึ่ม 18" = 1) OR (#"ปึ่ม 19" = 1) OR (#"ปึ่ม 20" = 1);
END_REGION
END_FUNCTION

FUNCTION "button start" : Void   // FC17, LAD
{ S7_Optimized_Access := 'TRUE' }
VERSION : 0.1
   VAR_OUTPUT
      Output : Bool;
   END_VAR
BEGIN

REGION Network 1
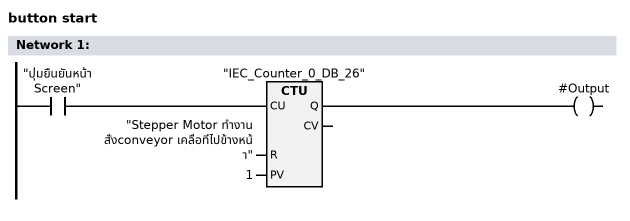
   "IEC_Counter_0_DB_26".CTU(CU := "ปุ่มยืนยันหน้า Screen",
                           R := "Stepper Motor ทำงาน สั่งconveyor เคลื่อที่ไปข้างหน้า",
                           PV := 1);
   #Output := "IEC_Counter_0_DB_26".Q;
END_REGION
END_FUNCTION

// folder: System_Out(เบิกจ่าย)/Gripperเบิกจ่าย

FUNCTION_BLOCK "Gripper_เบิกจ่าย"   // FB8, LAD
{ S7_Optimized_Access := 'TRUE' }
VERSION : 0.1
   VAR_TEMP   // added for the SCL form of the ladder/FBD networks
      _w1 : Bool;
   END_VAR
BEGIN

REGION Network 1
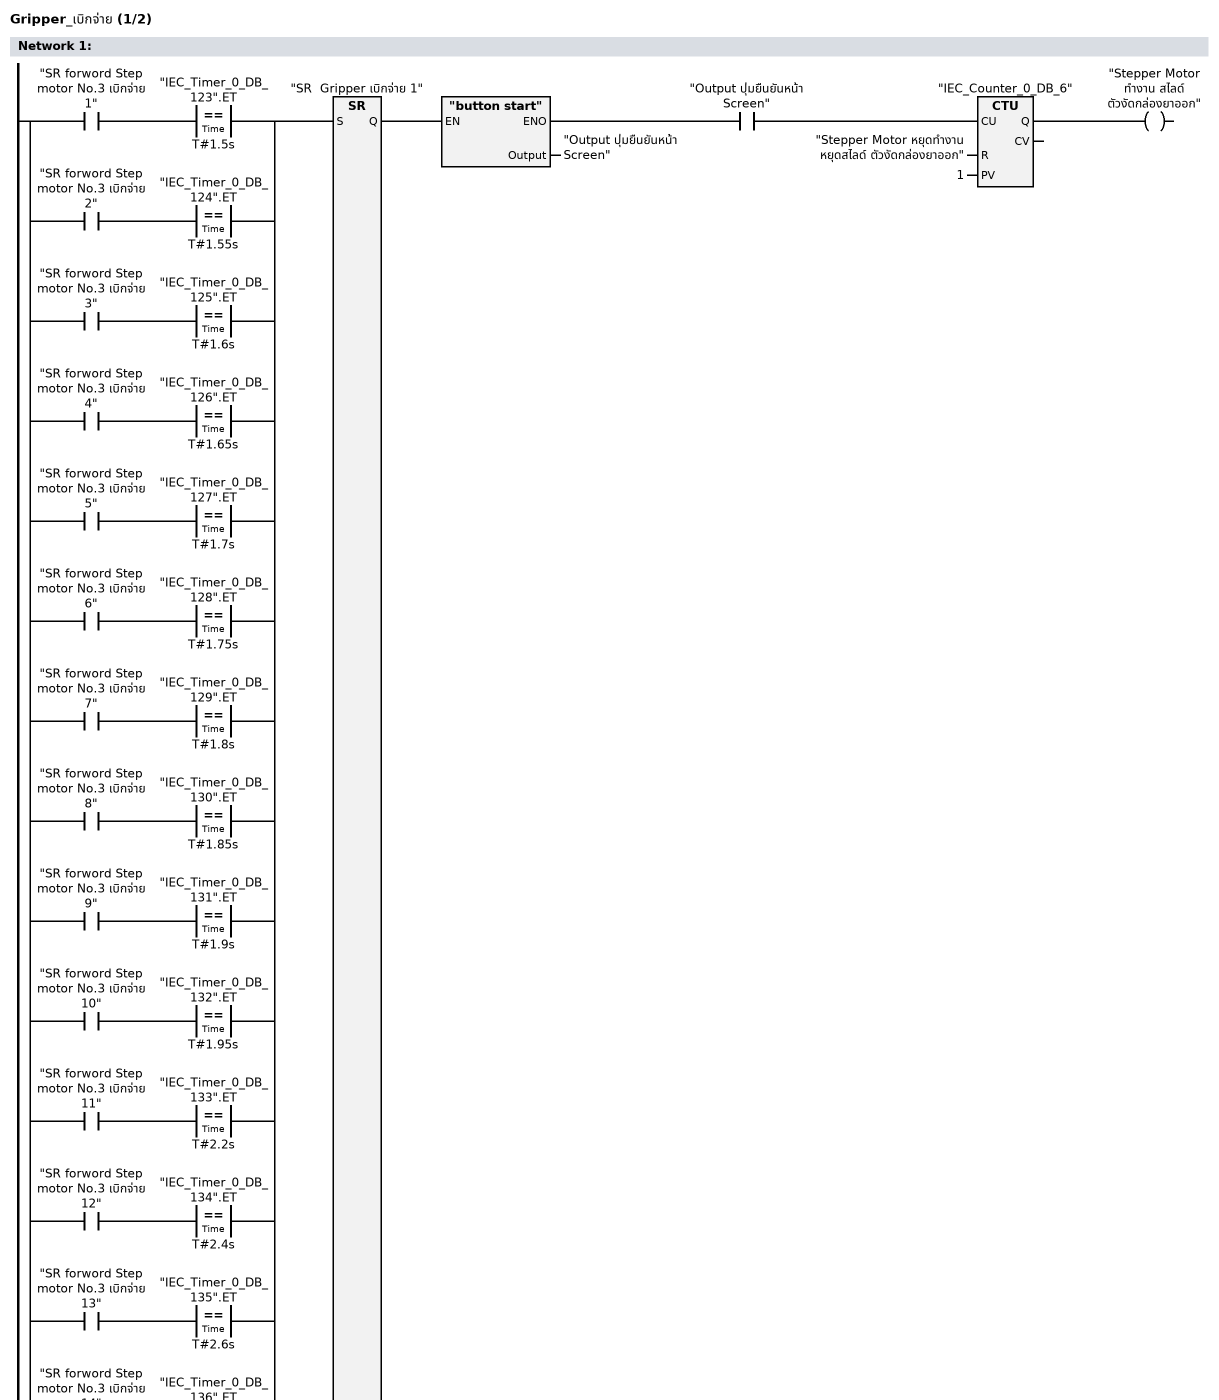
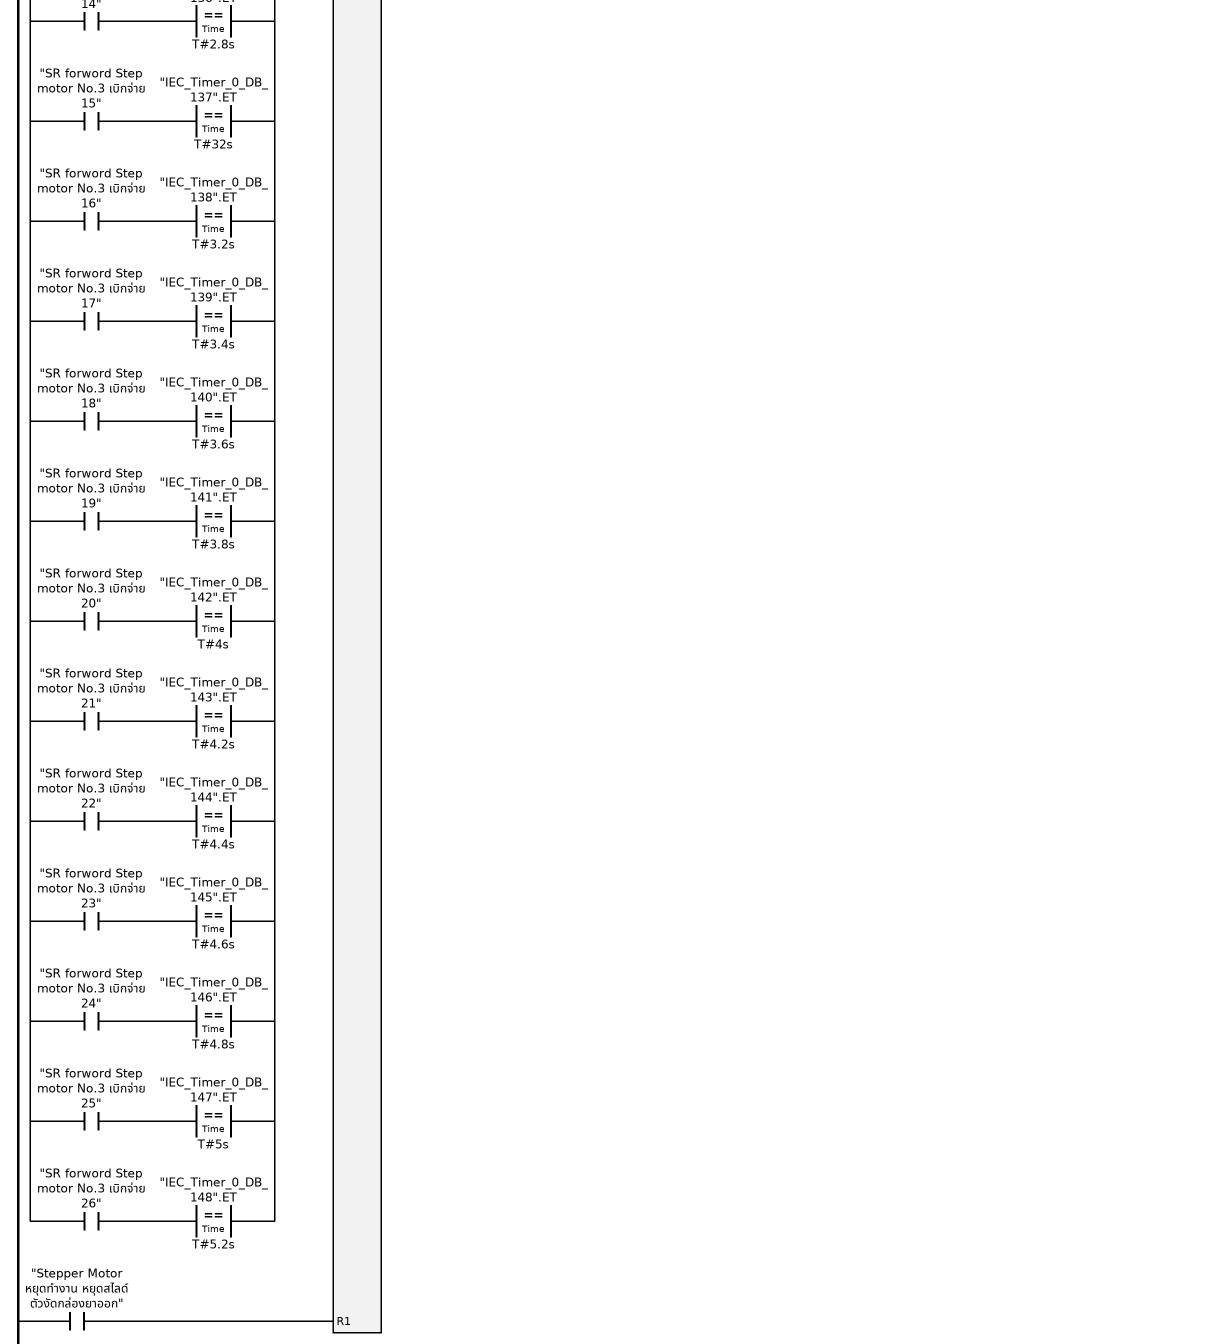
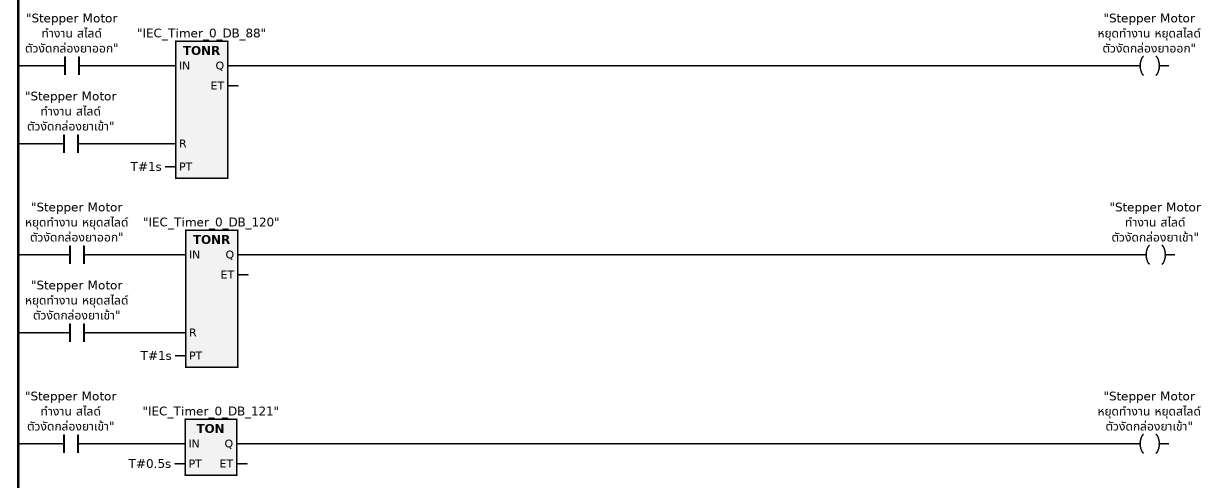
   IF ("SR forword Step motor No.3 เบิกจ่าย 1" AND ("IEC_Timer_0_DB_123".ET = T#1.5s)) OR ("SR forword Step motor No.3 เบิกจ่าย 2" AND ("IEC_Timer_0_DB_124".ET = T#1.55s)) OR ("SR forword Step motor No.3 เบิกจ่าย 3" AND ("IEC_Timer_0_DB_125".ET = T#1.6s)) OR ("SR forword Step motor No.3 เบิกจ่าย 4" AND ("IEC_Timer_0_DB_126".ET = T#1.65s)) OR ("SR forword Step motor No.3 เบิกจ่าย 5" AND ("IEC_Timer_0_DB_127".ET = T#1.7s)) OR ("SR forword Step motor No.3 เบิกจ่าย 6" AND ("IEC_Timer_0_DB_128".ET = T#1.75s)) OR ("SR forword Step motor No.3 เบิกจ่าย 7" AND ("IEC_Timer_0_DB_129".ET = T#1.8s)) OR ("SR forword Step motor No.3 เบิกจ่าย 8" AND ("IEC_Timer_0_DB_130".ET = T#1.85s)) OR ("SR forword Step motor No.3 เบิกจ่าย 9" AND ("IEC_Timer_0_DB_131".ET = T#1.9s)) OR ("SR forword Step motor No.3 เบิกจ่าย 10" AND ("IEC_Timer_0_DB_132".ET = T#1.95s)) OR ("SR forword Step motor No.3 เบิกจ่าย 11" AND ("IEC_Timer_0_DB_133".ET = T#2.2s)) OR ("SR forword Step motor No.3 เบิกจ่าย 12" AND ("IEC_Timer_0_DB_134".ET = T#2.4s)) OR ("SR forword Step motor No.3 เบิกจ่าย 13" AND ("IEC_Timer_0_DB_135".ET = T#2.6s)) OR ("SR forword Step motor No.3 เบิกจ่าย 14" AND ("IEC_Timer_0_DB_136".ET = T#2.8s)) OR ("SR forword Step motor No.3 เบิกจ่าย 15" AND ("IEC_Timer_0_DB_137".ET = T#32s)) OR ("SR forword Step motor No.3 เบิกจ่าย 16" AND ("IEC_Timer_0_DB_138".ET = T#3.2s)) OR ("SR forword Step motor No.3 เบิกจ่าย 17" AND ("IEC_Timer_0_DB_139".ET = T#3.4s)) OR ("SR forword Step motor No.3 เบิกจ่าย 18" AND ("IEC_Timer_0_DB_140".ET = T#3.6s)) OR ("SR forword Step motor No.3 เบิกจ่าย 19" AND ("IEC_Timer_0_DB_141".ET = T#3.8s)) OR ("SR forword Step motor No.3 เบิกจ่าย 20" AND ("IEC_Timer_0_DB_142".ET = T#4s)) OR ("SR forword Step motor No.3 เบิกจ่าย 21" AND ("IEC_Timer_0_DB_143".ET = T#4.2s)) OR ("SR forword Step motor No.3 เบิกจ่าย 22" AND ("IEC_Timer_0_DB_144".ET = T#4.4s)) OR ("SR forword Step motor No.3 เบิกจ่าย 23" AND ("IEC_Timer_0_DB_145".ET = T#4.6s)) OR ("SR forword Step motor No.3 เบิกจ่าย 24" AND ("IEC_Timer_0_DB_146".ET = T#4.8s)) OR ("SR forword Step motor No.3 เบิกจ่าย 25" AND ("IEC_Timer_0_DB_147".ET = T#5s)) OR ("SR forword Step motor No.3 เบิกจ่าย 26" AND ("IEC_Timer_0_DB_148".ET = T#5.2s)) THEN
       "SR  Gripper เบิกจ่าย 1" := TRUE;   // SR flip-flop
   END_IF;
   IF "Stepper Motor หยุดทำงาน หยุดสไลด์ ตัวงัดกล่องยาออก" THEN "SR  Gripper เบิกจ่าย 1" := FALSE; END_IF;
   "button start"(EN := "SR  Gripper เบิกจ่าย 1", Output => "Output ปุ่มยืนยันหน้า Screen", ENO => #_w1);
   "IEC_Counter_0_DB_6".CTU(CU := #_w1 AND "Output ปุ่มยืนยันหน้า Screen",
                           R := "Stepper Motor หยุดทำงาน หยุดสไลด์ ตัวงัดกล่องยาออก",
                           PV := 1);
   "Stepper Motor ทำงาน สไลด์ ตัวงัดกล่องยาออก" := "IEC_Counter_0_DB_6".Q;
   "IEC_Timer_0_DB_88".TONR(IN := "Stepper Motor ทำงาน สไลด์ ตัวงัดกล่องยาออก",
                           R := "Stepper Motor ทำงาน สไลด์ ตัวงัดกล่องยาเข้า",
                           PT := T#1s);
   "Stepper Motor หยุดทำงาน หยุดสไลด์ ตัวงัดกล่องยาออก" := "IEC_Timer_0_DB_88".Q;
   "IEC_Timer_0_DB_120".TONR(IN := "Stepper Motor หยุดทำงาน หยุดสไลด์ ตัวงัดกล่องยาออก",
                           R := "Stepper Motor หยุดทำงาน หยุดสไลด์ ตัวงัดกล่องยาเข้า",
                           PT := T#1s);
   "Stepper Motor ทำงาน สไลด์ ตัวงัดกล่องยาเข้า" := "IEC_Timer_0_DB_120".Q;
   "IEC_Timer_0_DB_121".TON(IN := "Stepper Motor ทำงาน สไลด์ ตัวงัดกล่องยาเข้า", PT := T#0.5s);
   "Stepper Motor หยุดทำงาน หยุดสไลด์ ตัวงัดกล่องยาเข้า" := "IEC_Timer_0_DB_121".Q;
END_REGION

REGION Network 2
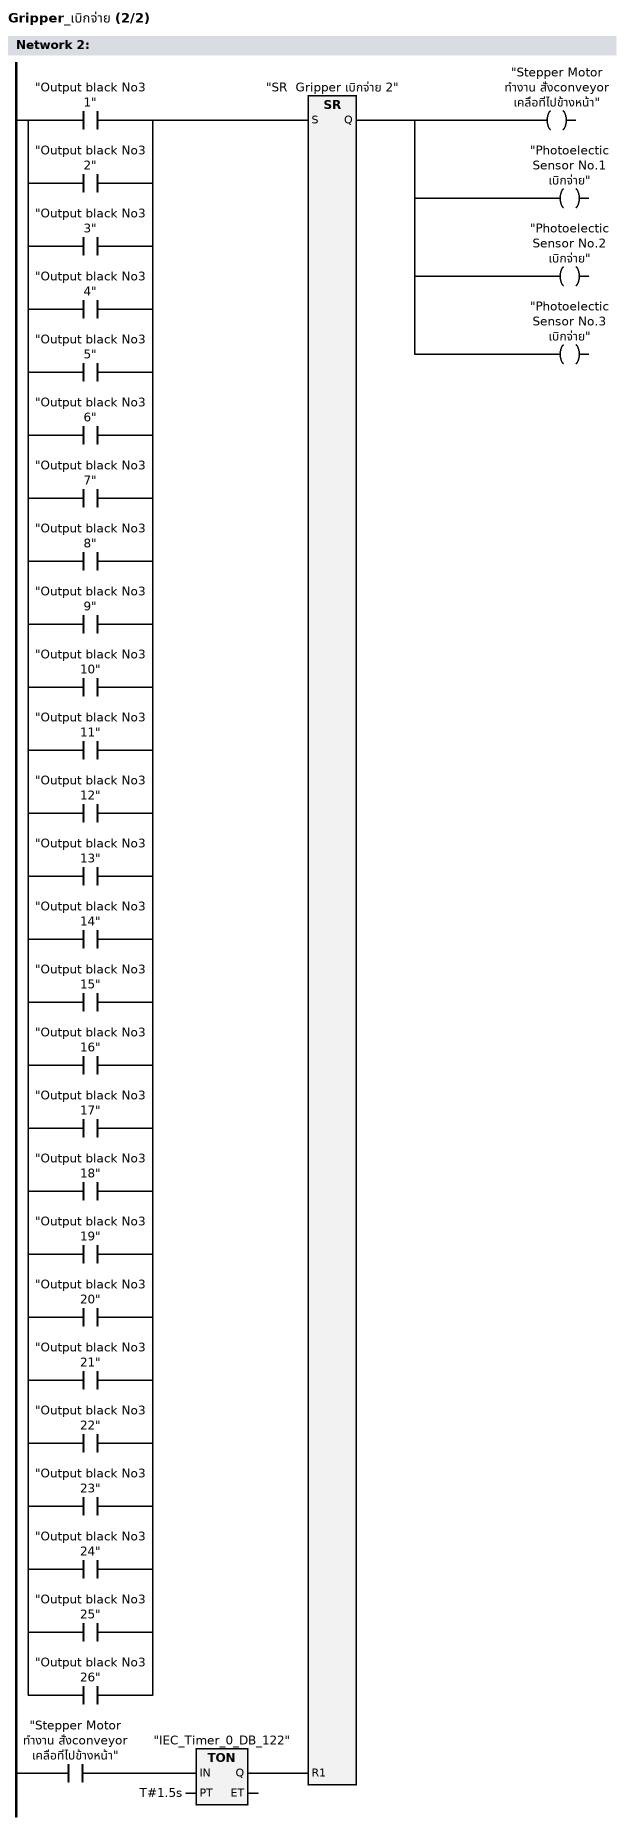
   "IEC_Timer_0_DB_122".TON(IN := "Stepper Motor ทำงาน สั่งconveyor เคลื่อที่ไปข้างหน้า", PT := T#1.5s);
   IF "Output black No3 1" OR "Output black No3 2" OR "Output black No3 3" OR "Output black No3 4" OR "Output black No3 5" OR "Output black No3 6" OR "Output black No3 7" OR "Output black No3 8" OR "Output black No3 9" OR "Output black No3 10" OR "Output black No3 11" OR "Output black No3 12" OR "Output black No3 13" OR "Output black No3 14" OR "Output black No3 15" OR "Output black No3 16" OR "Output black No3 17" OR "Output black No3 18" OR "Output black No3 19" OR "Output black No3 20" OR "Output black No3 21" OR "Output black No3 22" OR "Output black No3 23" OR "Output black No3 24" OR "Output black No3 25" OR "Output black No3 26" THEN
       "SR  Gripper เบิกจ่าย 2" := TRUE;   // SR flip-flop
   END_IF;
   IF "IEC_Timer_0_DB_122".Q THEN "SR  Gripper เบิกจ่าย 2" := FALSE; END_IF;
   "Stepper Motor ทำงาน สั่งconveyor เคลื่อที่ไปข้างหน้า" := "SR  Gripper เบิกจ่าย 2";
   "Photoelectic Sensor No.1 เบิกจ่าย" := "SR  Gripper เบิกจ่าย 2";
   "Photoelectic Sensor No.2 เบิกจ่าย" := "SR  Gripper เบิกจ่าย 2";
   "Photoelectic Sensor No.3 เบิกจ่าย" := "SR  Gripper เบิกจ่าย 2";
END_REGION
END_FUNCTION_BLOCK

FUNCTION "เวลาหลังจากเคลื่อนที่ถึงตำแหน่งเป้าหมาย (20)" : Void   // FC10, LAD
{ S7_Optimized_Access := 'TRUE' }
VERSION : 0.1
   VAR_INPUT
      "TONR 1" : Time;
      "Time 1" : Time;
      "TONR 2" : Time;
      "Time 2" : Time;
      "TONR 3" : Time;
      "Time 3" : Time;
      "TONR 4" : Time;
      "Time 4" : Time;
      "TONR 5" : Time;
      "Time 5" : Time;
      "TONR 6" : Time;
      "Time 6" : Time;
      "TONR 7" : Time;
      "Time 7" : Time;
      "TONR 8" : Time;
      "Time 8" : Time;
      "TONR 9" : Time;
      "Time 9" : Time;
      "TONR 10" : Time;
      "Time 10" : Time;
      "TONR 11" : Time;
      "Time 11" : Time;
      "TONR 12" : Time;
      "Time 12" : Time;
      "TONR 13" : Time;
      "Time 13" : Time;
      "TONR 14" : Time;
      "Time 14" : Time;
      "TONR 15" : Time;
      "Time 15" : Time;
      "TONR 16" : Time;
      "Time 16" : Time;
      "TONR 17" : Time;
      "Time 17" : Time;
      "TONR 18" : Time;
      "Time 18" : Time;
      "TONR 19" : Time;
      "Time 19" : Time;
      "TONR 20" : Time;
      "Time 20" : Time;
      "TONR 21" : Time;
      "Time 21" : Time;
      "TONR 22" : Time;
      "Time 22" : Time;
      "TONR 23" : Time;
      "Time 23" : Time;
      "TONR 24" : Time;
      "Time 24" : Time;
      "TONR 25" : Time;
      "Time 25" : Time;
      "TONR 26" : Time;
      "Time 26" : Time;
   END_VAR
   VAR_OUTPUT
      "Output Time" : Bool;
   END_VAR
BEGIN

REGION Network 1
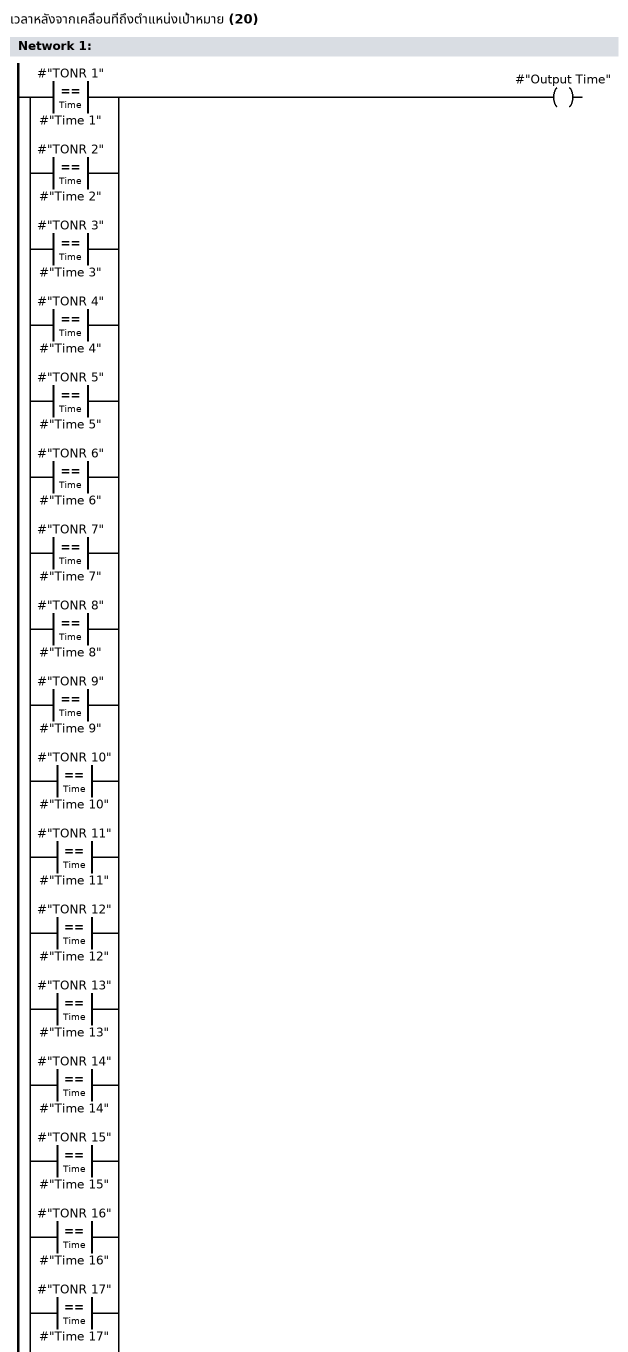
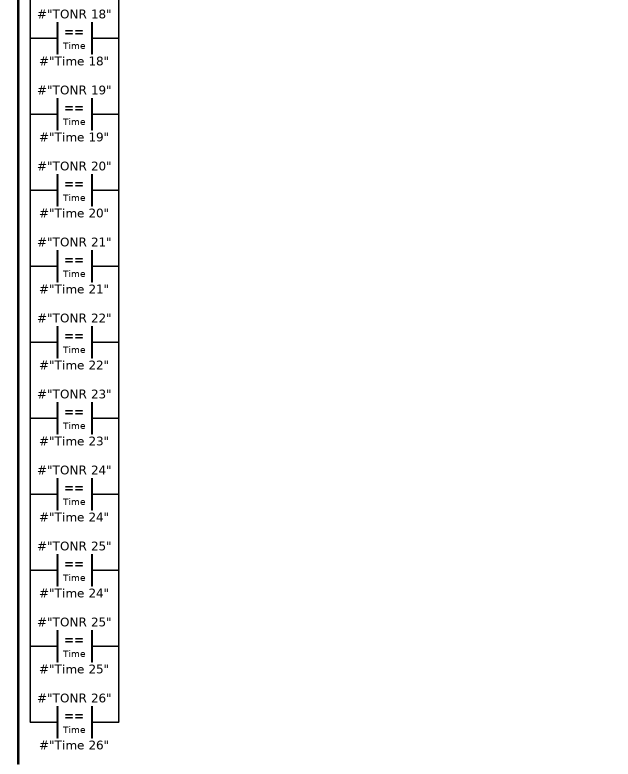
   RUNG wire#powerrail
      { S7_Templates := "SrcType := Time" } EQ_Contact(in1 := #"TONR 1", in2 := #"Time 1")
      wire#w1
      Coil( #"Output Time" )
   END_RUNG
   RUNG wire#powerrail
      { S7_Templates := "SrcType := Time" } EQ_Contact(in1 := #"TONR 2", in2 := #"Time 2")
   END_RUNG wire#w1
   RUNG wire#powerrail
      { S7_Templates := "SrcType := Time" } EQ_Contact(in1 := #"TONR 3", in2 := #"Time 3")
   END_RUNG wire#w1
   RUNG wire#powerrail
      { S7_Templates := "SrcType := Time" } EQ_Contact(in1 := #"TONR 4", in2 := #"Time 4")
   END_RUNG wire#w1
   RUNG wire#powerrail
      { S7_Templates := "SrcType := Time" } EQ_Contact(in1 := #"TONR 5", in2 := #"Time 5")
   END_RUNG wire#w1
   RUNG wire#powerrail
      { S7_Templates := "SrcType := Time" } EQ_Contact(in1 := #"TONR 6", in2 := #"Time 6")
   END_RUNG wire#w1
   RUNG wire#powerrail
      { S7_Templates := "SrcType := Time" } EQ_Contact(in1 := #"TONR 7", in2 := #"Time 7")
   END_RUNG wire#w1
   RUNG wire#powerrail
      { S7_Templates := "SrcType := Time" } EQ_Contact(in1 := #"TONR 8", in2 := #"Time 8")
   END_RUNG wire#w1
   RUNG wire#powerrail
      { S7_Templates := "SrcType := Time" } EQ_Contact(in1 := #"TONR 9", in2 := #"Time 9")
   END_RUNG wire#w1
   RUNG wire#powerrail
      { S7_Templates := "SrcType := Time" } EQ_Contact(in1 := #"TONR 10", in2 := #"Time 10")
   END_RUNG wire#w1
   RUNG wire#powerrail
      { S7_Templates := "SrcType := Time" } EQ_Contact(in1 := #"TONR 11", in2 := #"Time 11")
   END_RUNG wire#w1
   RUNG wire#powerrail
      { S7_Templates := "SrcType := Time" } EQ_Contact(in1 := #"TONR 12", in2 := #"Time 12")
   END_RUNG wire#w1
   RUNG wire#powerrail
      { S7_Templates := "SrcType := Time" } EQ_Contact(in1 := #"TONR 13", in2 := #"Time 13")
   END_RUNG wire#w1
   RUNG wire#powerrail
      { S7_Templates := "SrcType := Time" } EQ_Contact(in1 := #"TONR 14", in2 := #"Time 14")
   END_RUNG wire#w1
   RUNG wire#powerrail
      { S7_Templates := "SrcType := Time" } EQ_Contact(in1 := #"TONR 15", in2 := #"Time 15")
   END_RUNG wire#w1
   RUNG wire#powerrail
      { S7_Templates := "SrcType := Time" } EQ_Contact(in1 := #"TONR 16", in2 := #"Time 16")
   END_RUNG wire#w1
   RUNG wire#powerrail
      { S7_Templates := "SrcType := Time" } EQ_Contact(in1 := #"TONR 17", in2 := #"Time 17")
   END_RUNG wire#w1
   RUNG wire#powerrail
      { S7_Templates := "SrcType := Time" } EQ_Contact(in1 := #"TONR 18", in2 := #"Time 18")
   END_RUNG wire#w1
   RUNG wire#powerrail
      { S7_Templates := "SrcType := Time" } EQ_Contact(in1 := #"TONR 19", in2 := #"Time 19")
   END_RUNG wire#w1
   RUNG wire#powerrail
      { S7_Templates := "SrcType := Time" } EQ_Contact(in1 := #"TONR 20", in2 := #"Time 20")
   END_RUNG wire#w1
   RUNG wire#powerrail
      { S7_Templates := "SrcType := Time" } EQ_Contact(in1 := #"TONR 21", in2 := #"Time 21")
   END_RUNG wire#w1
   RUNG wire#powerrail
      { S7_Templates := "SrcType := Time" } EQ_Contact(in1 := #"TONR 22", in2 := #"Time 22")
   END_RUNG wire#w1
   RUNG wire#powerrail
      { S7_Templates := "SrcType := Time" } EQ_Contact(in1 := #"TONR 23", in2 := #"Time 23")
   END_RUNG wire#w1
   RUNG wire#powerrail
      { S7_Templates := "SrcType := Time" } EQ_Contact(in1 := #"TONR 24", in2 := #"Time 24")
   END_RUNG wire#w1
   RUNG wire#powerrail
      { S7_Templates := "SrcType := Time" } EQ_Contact(in1 := #"TONR 25", in2 := #"Time 24")
   END_RUNG wire#w1
   RUNG wire#powerrail
      { S7_Templates := "SrcType := Time" } EQ_Contact(in1 := #"TONR 25", in2 := #"Time 25")
   END_RUNG wire#w1
   RUNG wire#powerrail
      { S7_Templates := "SrcType := Time" } EQ_Contact(in1 := #"TONR 26", in2 := #"Time 26")
   END_RUNG wire#w1
   // the same network as SCL:
   #"Output Time" := (#"TONR 1" = #"Time 1") OR (#"TONR 2" = #"Time 2") OR (#"TONR 3" = #"Time 3") OR (#"TONR 4" = #"Time 4") OR (#"TONR 5" = #"Time 5") OR (#"TONR 6" = #"Time 6") OR (#"TONR 7" = #"Time 7") OR (#"TONR 8" = #"Time 8") OR (#"TONR 9" = #"Time 9") OR (#"TONR 10" = #"Time 10") OR (#"TONR 11" = #"Time 11") OR (#"TONR 12" = #"Time 12") OR (#"TONR 13" = #"Time 13") OR (#"TONR 14" = #"Time 14") OR (#"TONR 15" = #"Time 15") OR (#"TONR 16" = #"Time 16") OR (#"TONR 17" = #"Time 17") OR (#"TONR 18" = #"Time 18") OR (#"TONR 19" = #"Time 19") OR (#"TONR 20" = #"Time 20") OR (#"TONR 21" = #"Time 21") OR (#"TONR 22" = #"Time 22") OR (#"TONR 23" = #"Time 23") OR (#"TONR 24" = #"Time 24") OR (#"TONR 25" = #"Time 24") OR (#"TONR 25" = #"Time 25") OR (#"TONR 26" = #"Time 26");
END_REGION
END_FUNCTION

FUNCTION "Test-----1" : Void   // FC12, LAD
{ S7_Optimized_Access := 'TRUE' }
VERSION : 0.1
   VAR_INPUT
      "TONR 1" : Time;
      "Time 1" : Time;
      "TONR 2" : Time;
      "Time 2" : Time;
      "TONR 3" : Time;
      "Time 3" : Time;
      "TONR 4" : Time;
      "Time 4" : Time;
      "TONR 5" : Time;
      "Time 5" : Time;
      "TONR 6" : Time;
      "Time 6" : Time;
      "TONR 7" : Time;
      "Time 7" : Time;
      "TONR 8" : Time;
      "Time 8" : Time;
      "TONR 9" : Time;
      "Time 9" : Time;
      "TONR 10" : Time;
      "Time 10" : Time;
      "TONR 11" : Time;
      "Time 11" : Time;
      "TONR 12" : Time;
      "Time 12" : Time;
      "TONR 13" : Time;
      "Time 13" : Time;
      "TONR 14" : Time;
      "Time 14" : Time;
      "TONR 15" : Time;
      "Time 15" : Time;
      "TONR 16" : Time;
      "Time 16" : Time;
      "TONR 17" : Time;
      "Time 17" : Time;
      "TONR 18" : Time;
      "Time 18" : Time;
      "TONR 19" : Time;
      "Time 19" : Time;
      "TONR 20" : Time;
      "Time 20" : Time;
   END_VAR
   VAR_OUTPUT
      "Output Time" : Bool;
   END_VAR
BEGIN

REGION Network 1
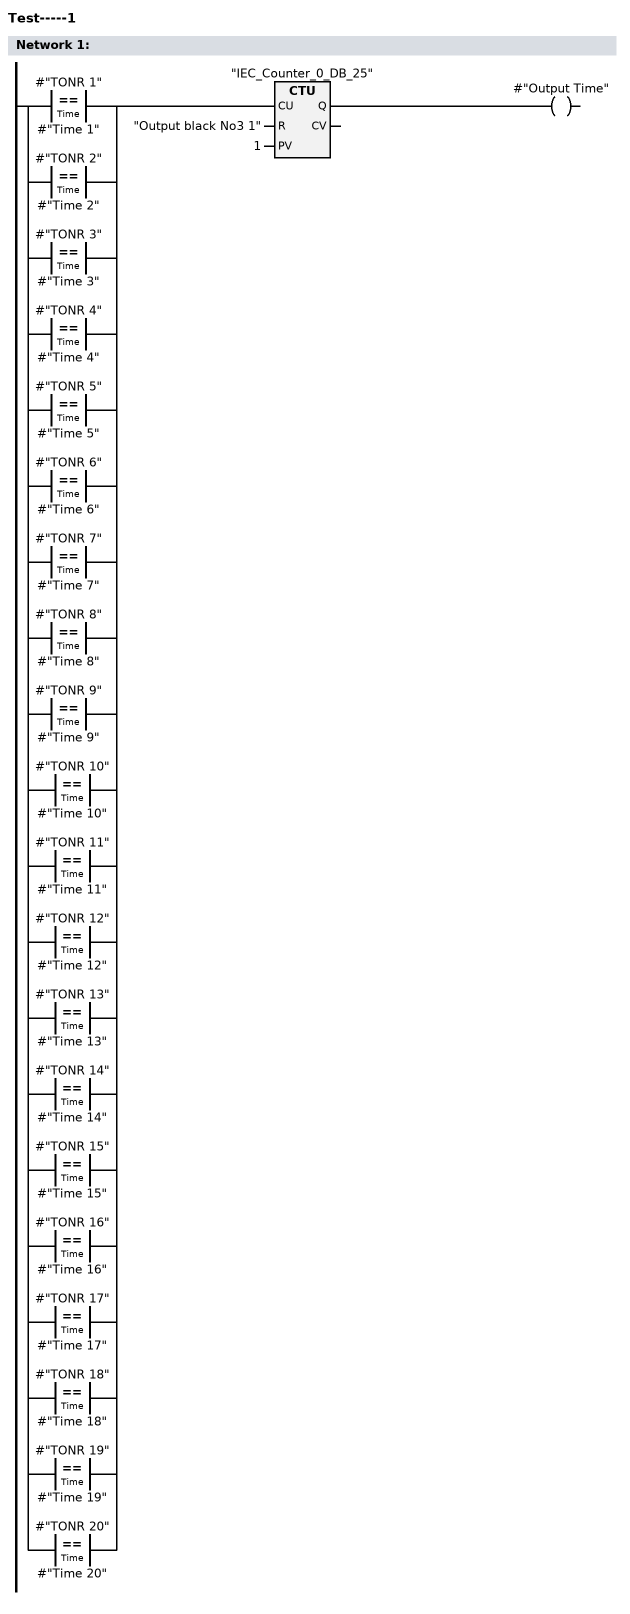
   "IEC_Counter_0_DB_25".CTU(CU := (#"TONR 1" = #"Time 1") OR (#"TONR 2" = #"Time 2") OR (#"TONR 3" = #"Time 3") OR (#"TONR 4" = #"Time 4") OR (#"TONR 5" = #"Time 5") OR (#"TONR 6" = #"Time 6") OR (#"TONR 7" = #"Time 7") OR (#"TONR 8" = #"Time 8") OR (#"TONR 9" = #"Time 9") OR (#"TONR 10" = #"Time 10") OR (#"TONR 11" = #"Time 11") OR (#"TONR 12" = #"Time 12") OR (#"TONR 13" = #"Time 13") OR (#"TONR 14" = #"Time 14") OR (#"TONR 15" = #"Time 15") OR (#"TONR 16" = #"Time 16") OR (#"TONR 17" = #"Time 17") OR (#"TONR 18" = #"Time 18") OR (#"TONR 19" = #"Time 19") OR (#"TONR 20" = #"Time 20"),
                           R := "Output black No3 1",
                           PV := 1);
   #"Output Time" := "IEC_Counter_0_DB_25".Q;
END_REGION
END_FUNCTION

// folder: System_Out(เบิกจ่าย)/Step motor No.1,No.2(เบิกจาย)

FUNCTION_BLOCK "Step motor ขึ่น-ลง ตามแกน y No.1,No.2_Forword(เบิกจ่าย)"   // FB5, LAD
{ S7_Optimized_Access := 'TRUE' }
VERSION : 0.1
   VAR_INPUT
      "TIME ที่ใช้ไป BOX.1-BOX.26 เบิกจ่าย" : Time;
      "TIME ที่ใช้ไป BOX.27-BOX.52 เบิกจ่าย" : Time;
      "TIME ที่ใช้ไป BOX.53-BOX.78เบิกจ่าย" : Time;
      "TIME ที่ใช้ไป BOX.79-BOX.104เบิกจ่าย" : Time;
      "TIME ที่ใช้ไป BOX.105-BOX.130เบิกจ่าย" : Time;
      "TIME ที่ใช้ไป BOX.131-BOX.156เบิกจ่าย" : Time;
      "TIME ที่ใช้ไป BOX.157-BOX.182เบิกจ่าย" : Time;
      "TIME ที่ใช้ไป BOX.183-BOX.208เบิกจ่าย" : Time;
      "TIME ที่ใช้ไป BOX.209-BOX.234เบิกจ่าย" : Time;
      "TIME ที่ใช้ไป BOX.235-BOX.260เบิกจ่าย" : Time;
      "TIME ที่ใช้ไป BOX.261-BOX.286เบิกจ่าย" : Time;
      "TIME ที่ใช้ไป BOX.287-BOX.312เบิกจ่าย" : Time;
      "TIME ที่ใช้ไป BOX.313-BOX.338เบิกจ่าย" : Time;
      "TIME ที่ใช้ไป BOX.339-BOX.364เบิกจ่าย" : Time;
      "TIME ที่ใช้ไป BOX.365-BOX.390เบิกจ่าย" : Time;
      "TIME ที่ใช้ไป BOX.391-BOX.416เบิกจ่าย" : Time;
      "TIME ที่ใช้ไป BOX.417-BOX.442เบิกจ่าย" : Time;
      "TIME ที่ใช้ไป BOX.443-BOX.468เบิกจ่าย" : Time;
      "TIME ที่ใช้ไป BOX.469-BOX.494เบิกจ่าย" : Time;
      "TIME ที่ใช้ไป BOX.495-BOX.520เบิกจ่าย" : Time;
   END_VAR
   VAR_IN_OUT
      "Stepper Motor  ทำงาน" : Bool;
   END_VAR
   VAR_TEMP   // added for the SCL form of the ladder/FBD networks
      _w1 : Bool;
      _w2 : Bool;
      _w3 : Bool;
      _w4 : Bool;
      _w5 : Bool;
      _w6 : Bool;
      _w7 : Bool;
      _w8 : Bool;
      _w9 : Bool;
      _w10 : Bool;
      _w11 : Bool;
      _w12 : Bool;
      _w13 : Bool;
      _w14 : Bool;
      _w15 : Bool;
      _w16 : Bool;
      _w17 : Bool;
      _w18 : Bool;
      _w19 : Bool;
      _w20 : Bool;
      _w21 : Bool;
      _w22 : Bool;
      _w23 : Bool;
      _w24 : Bool;
      _w25 : Bool;
      _w26 : Bool;
      _w27 : Bool;
      _w28 : Bool;
      _w29 : Bool;
      _w30 : Bool;
      _w31 : Bool;
      _w32 : Bool;
      _w33 : Bool;
      _w34 : Bool;
      _w35 : Bool;
      _w36 : Bool;
      _w37 : Bool;
      _w38 : Bool;
      _w39 : Bool;
      _w40 : Bool;
      _w41 : Bool;
      _w42 : Bool;
      _w43 : Bool;
      _w44 : Bool;
      _w45 : Bool;
      _w46 : Bool;
      _w47 : Bool;
      _w48 : Bool;
      _w49 : Bool;
      _w50 : Bool;
      _w51 : Bool;
      _w52 : Bool;
      _w53 : Bool;
      _w54 : Bool;
      _w55 : Bool;
      _w56 : Bool;
      _w57 : Bool;
      _w58 : Bool;
      _w59 : Bool;
   END_VAR
BEGIN

REGION Network 1
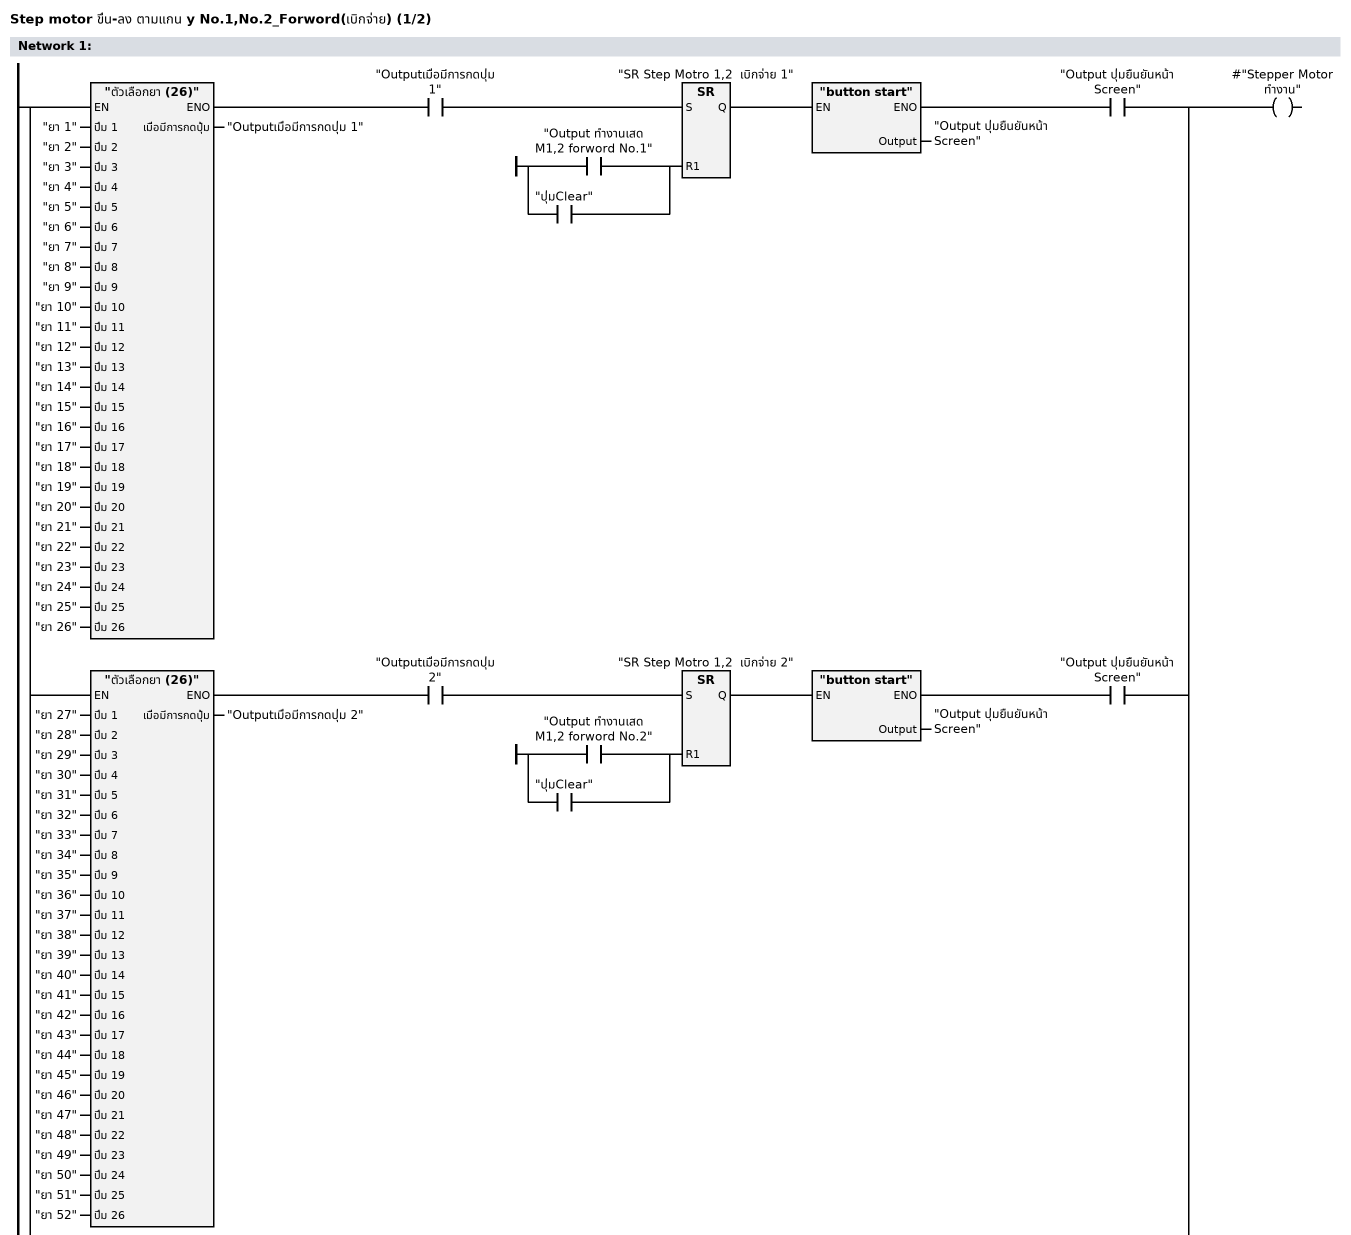
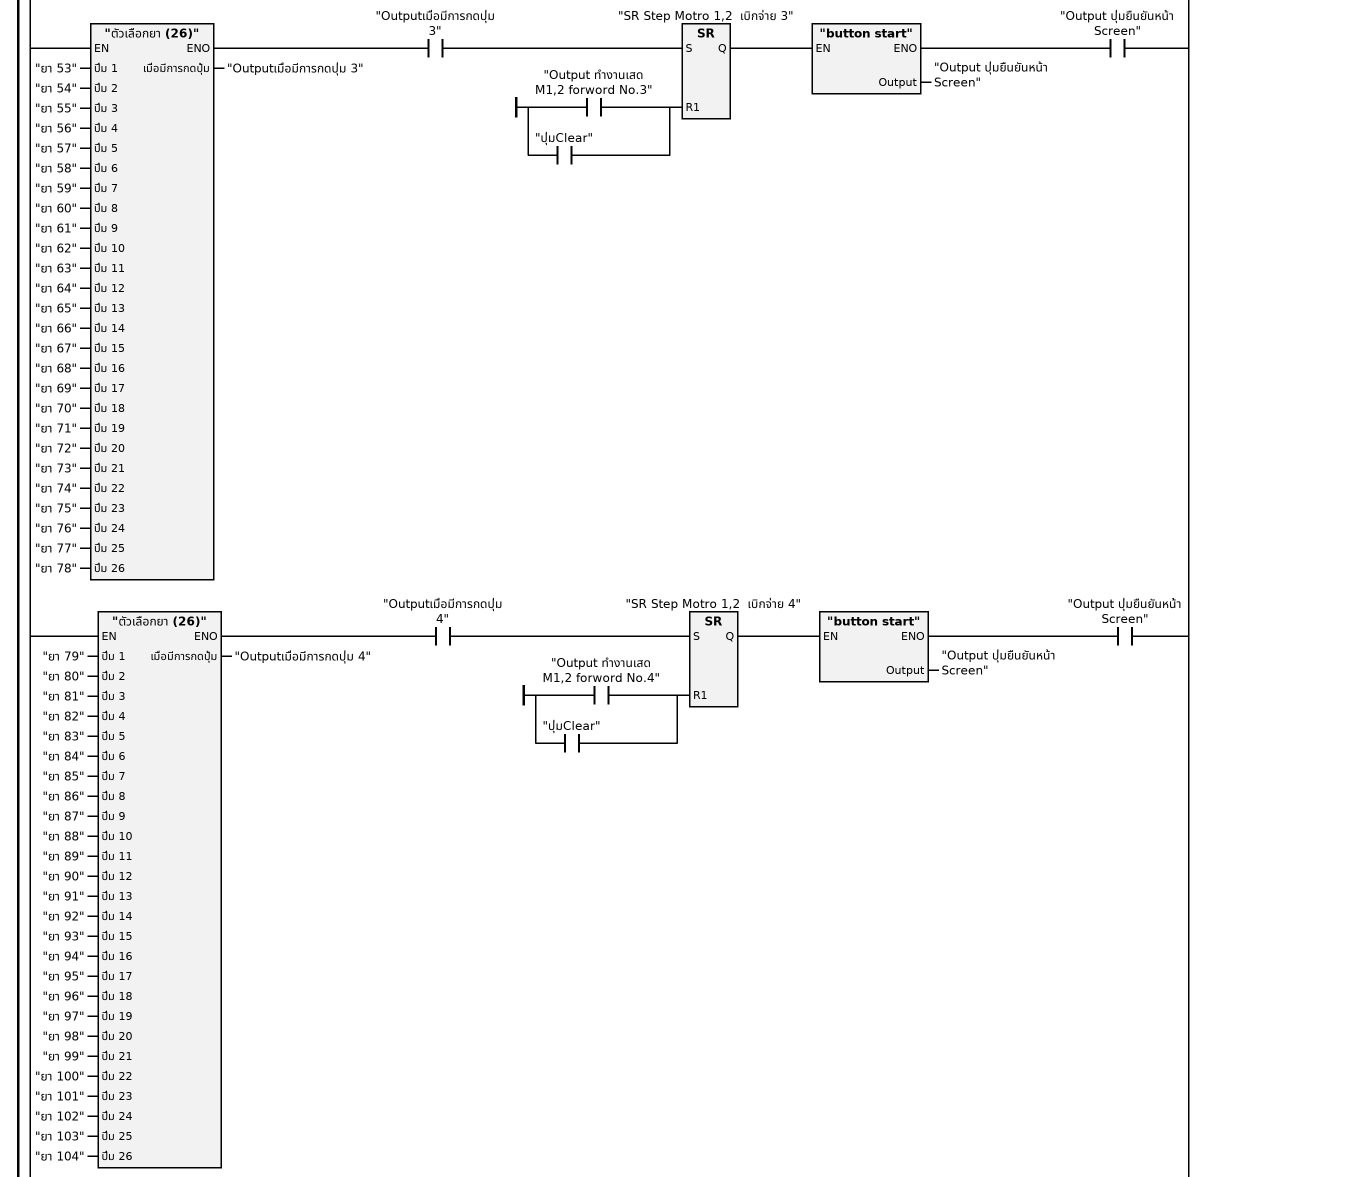
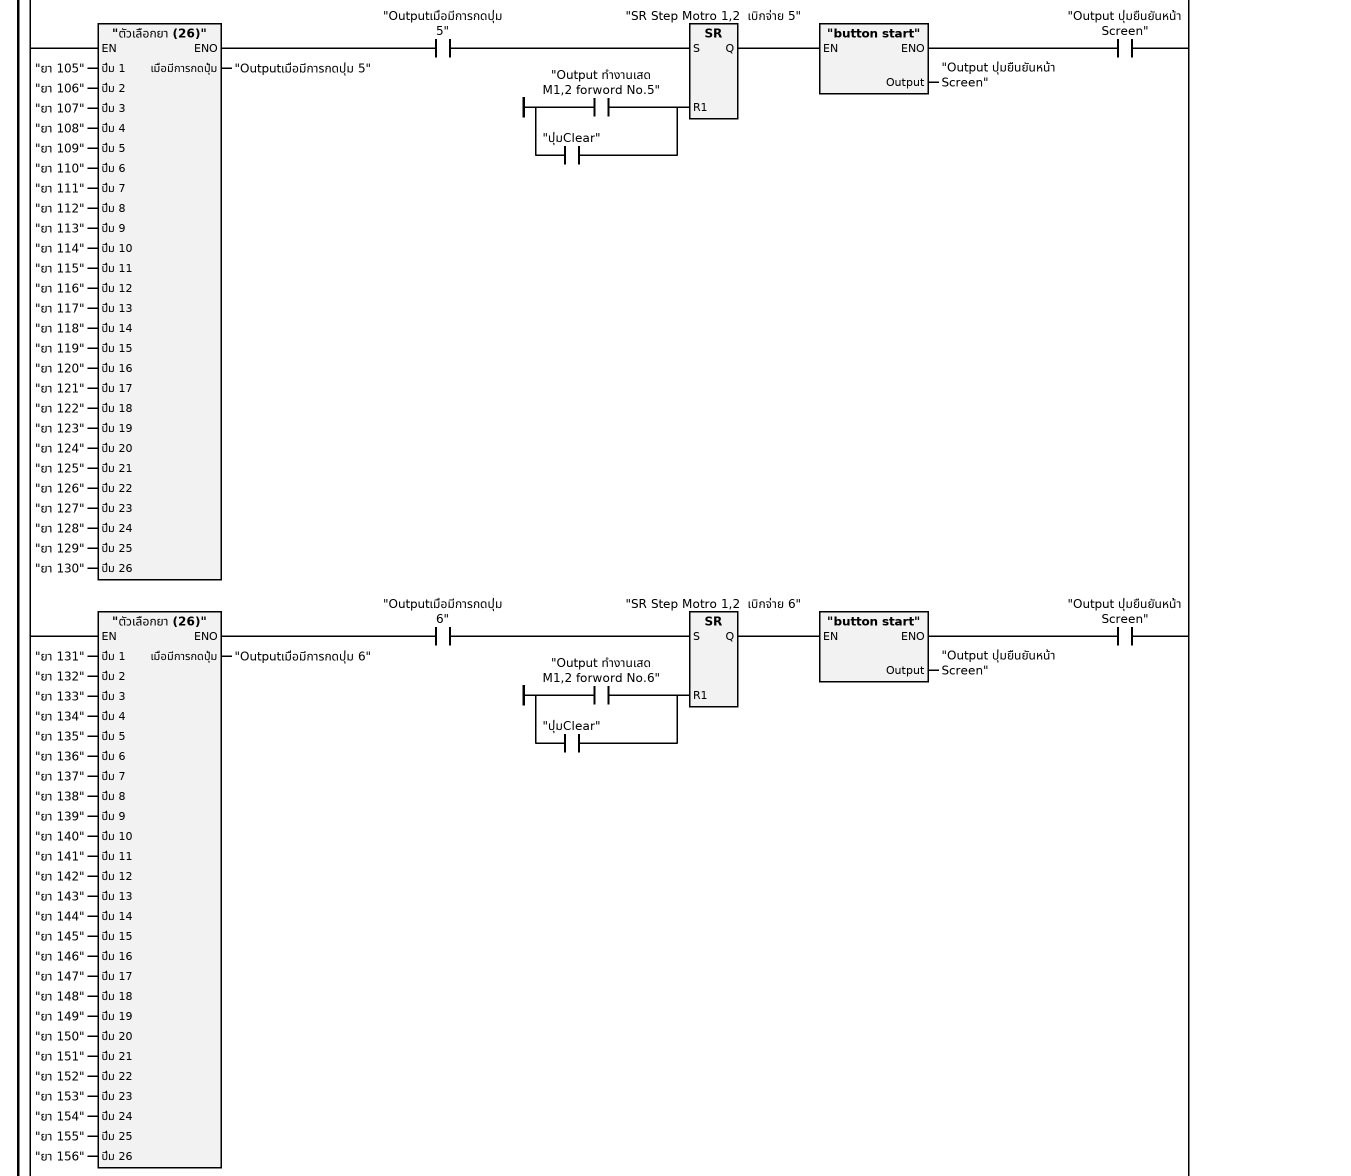
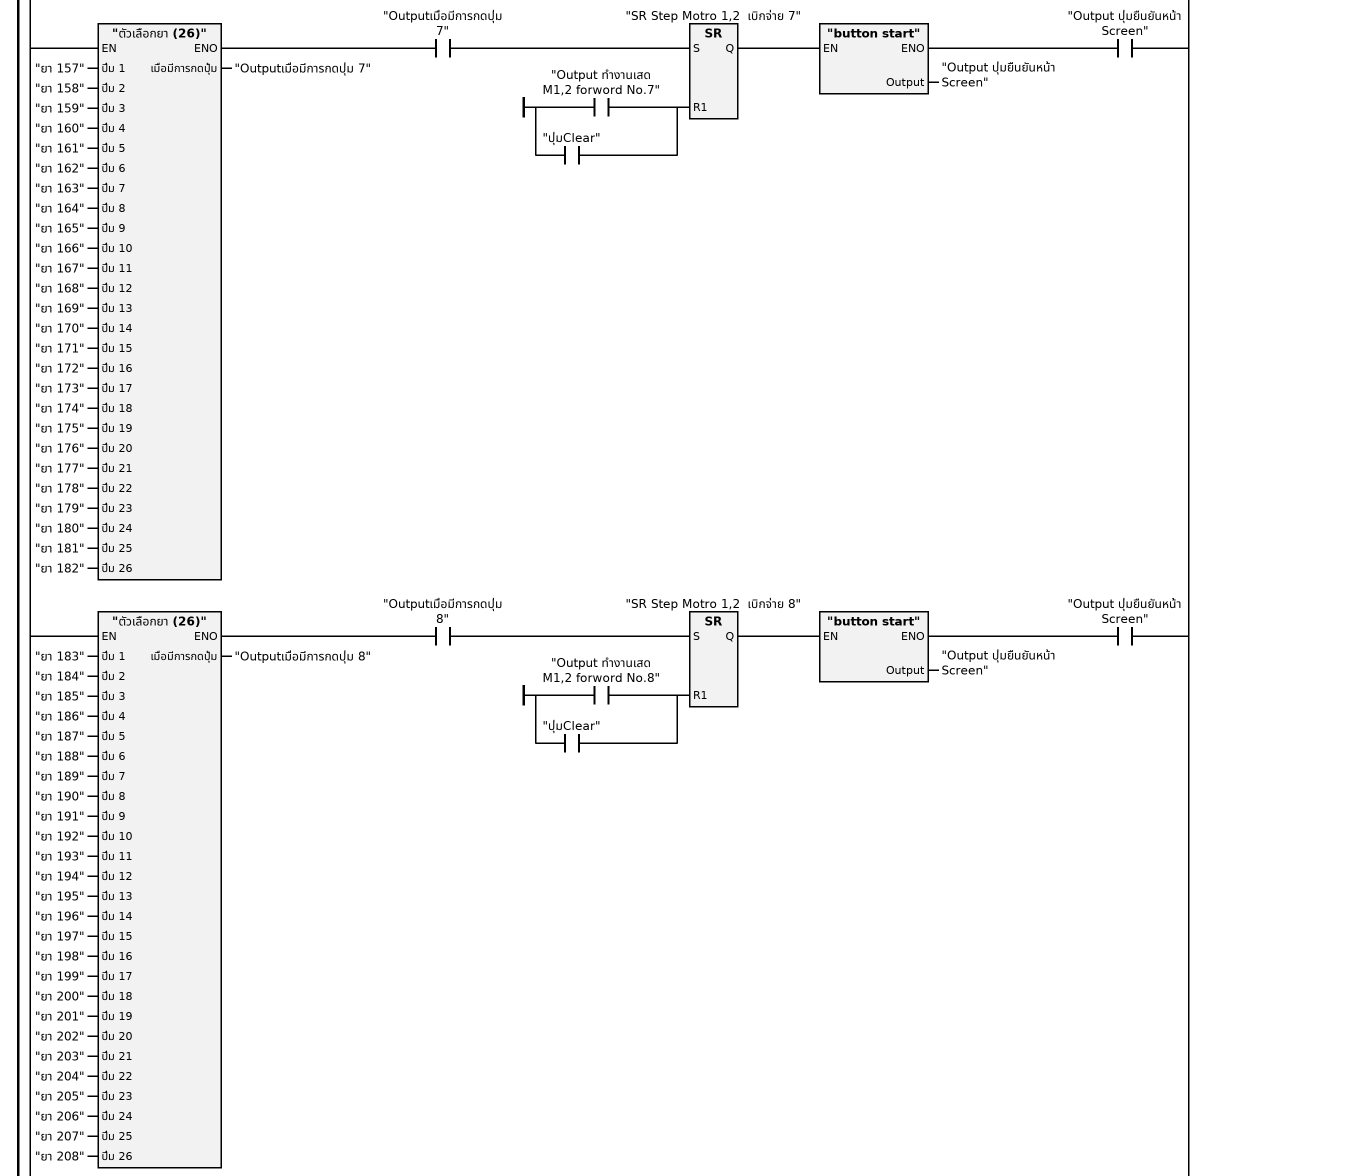
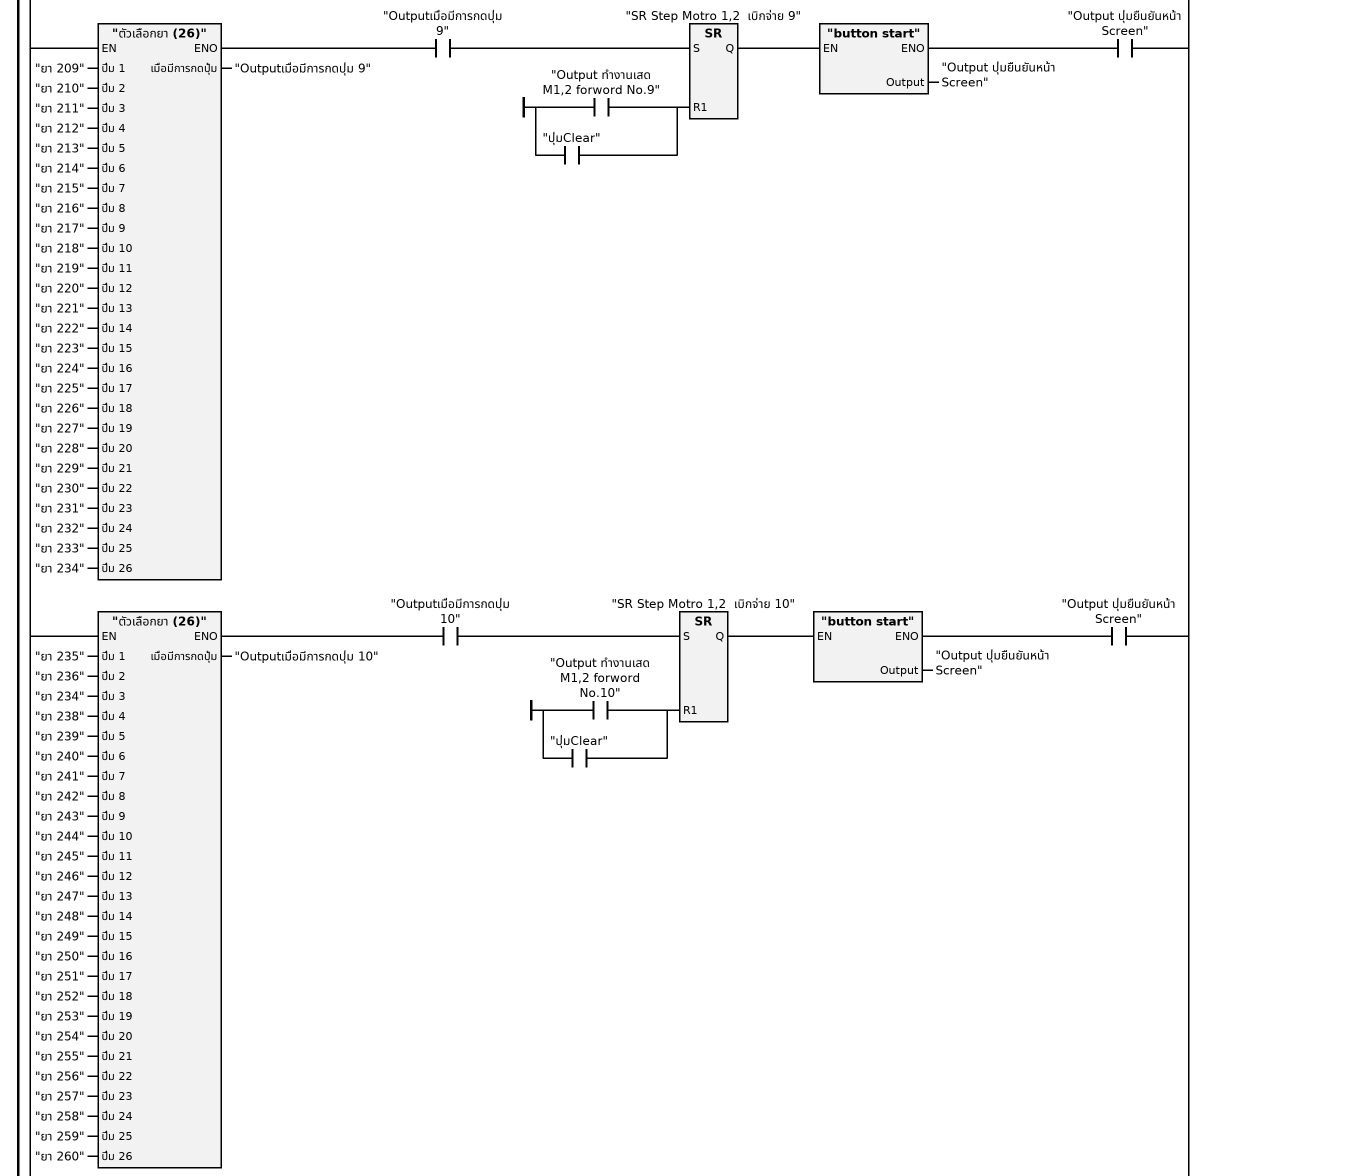
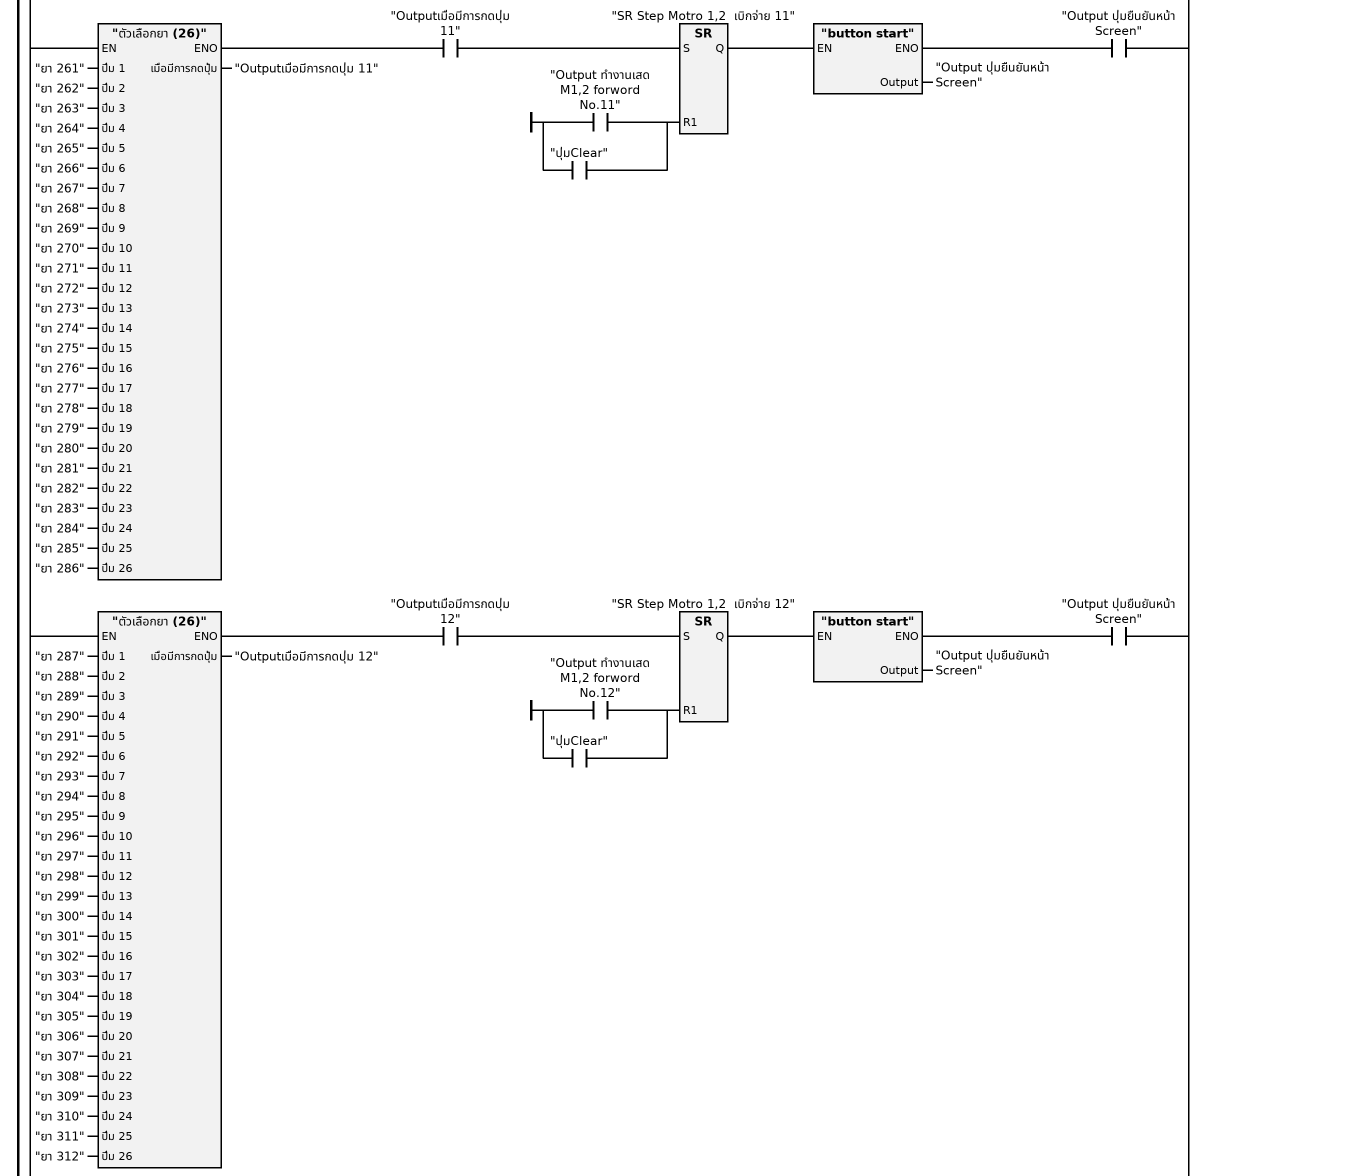
